   //Copy data
   FOR #i := 1 TO 9 DO
       #j := "HMI_OrderTable".StartRow + #i;
       "HMI_OrderTable".Index[#i] := #j;
       "HMI_OrderTable".OrderTable[#i] := #System.OrderTable[#j];
       //Color State
       IF "HMI_OrderTable".OrderTable[#i].Status = 'Queued' THEN
           "HMI_OrderTable".State[#i] := 1;
       ELSIF "HMI_OrderTable".OrderTable[#i].Status = 'Running' THEN
           "HMI_OrderTable".State[#i] := 2;
       ELSIF "HMI_OrderTable".OrderTable[#i].Status = 'Completed' THEN
           "HMI_OrderTable".State[#i] := 3;
       ELSIF "HMI_OrderTable".OrderTable[#i].Status = 'Error' THEN
           "HMI_OrderTable".State[#i] := 4;
       ELSIF "HMI_OrderTable".OrderTable[#i].Status = 'Paused' THEN
           "HMI_OrderTable".State[#i] := 5;
       ELSIF "HMI_OrderTable".OrderTable[#i].Status = 'Canceled' THEN
           "HMI_OrderTable".State[#i] := 6;
       ELSIF "HMI_OrderTable".OrderTable[#i].Status = 'Error\Cancel' THEN
           "HMI_OrderTable".State[#i] := 7;
       ELSE
           "HMI_OrderTable".State[#i] := 0;
       END_IF;
   END_FOR;

   IF NOT "HMI_OrderTable".PlacingNewOrder THEN
       "HMI_OrderTable".Device := 0;
   END_IF;

   //Error PopUp Window
   IF "HMI_OrderTable".PopUp_ErrorWindow_Active AND NOT "HMI_OrderTable".PlacingNewOrder THEN
       "HMI_OrderTable".OrderTable[0] := "HMI_OrderTable".OrderTable["HMI_OrderTable".PopUp_Index];
       IF "HMI_OrderTable".OrderTable[0].Status = 'Error' THEN
           "HMI_OrderTable".State[0] := 4;
       ELSIF "HMI_OrderTable".OrderTable[0].Status = 'Error\Cancel' THEN
           "HMI_OrderTable".State[0] := 7;
       ELSE
           "HMI_OrderTable".State[0] := 0;
       END_IF;
   ELSIF NOT "HMI_OrderTable".PopUp_ErrorWindow_Active AND NOT "HMI_OrderTable".PlacingNewOrder THEN
       "HMI_OrderTable".OrderTable[0] := #EmptyOrder;
   END_IF;

   REGION Testing area
       IF ("HMI_Box_Connected_1" = #System.Id OR ("HMI_Box_Connected_1" >= (#System.Id * 10) + 1 AND "HMI_Box_Connected_1" <= (#System.Id * 10) + 8)) OR
           ("HMI_Box_Connected_2" = #System.Id OR ("HMI_Box_Connected_1" >= (#System.Id * 10) + 1 AND "HMI_Box_Connected_1" <= (#System.Id * 10) + 8))
       THEN
           #System_Busy := TRUE;
       ELSE
           #System_Busy := FALSE;
           IF "Comissioning_Var" THEN
           //Visibilities
           //Running in auto mode
           IF #Auto_Test.Running AND NOT #Auto_Test.Manual AND NOT #Auto_Test.Pause THEN
               "OrderTable_HMI"."Start Test Visibility" := FALSE;
               "OrderTable_HMI"."Stop Test Visibility" := TRUE;
               "OrderTable_HMI"."Pause Test Visibility" := TRUE;
               "OrderTable_HMI"."Resume Visibility" := FALSE;
               "OrderTable_HMI"."Clear Table Visibility" := FALSE;
               "OrderTable_HMI"."Manual order Visibility" := FALSE;
               //Running and paused
           ELSIF #Auto_Test.Running AND #Auto_Test.Pause AND NOT #Auto_Test.Manual THEN
               "OrderTable_HMI"."Start Test Visibility" := FALSE;
               "OrderTable_HMI"."Stop Test Visibility" := TRUE;
               "OrderTable_HMI"."Pause Test Visibility" := FALSE;
               "OrderTable_HMI"."Resume Visibility" := TRUE;
               "OrderTable_HMI"."Clear Table Visibility" := FALSE;
               "OrderTable_HMI"."Manual order Visibility" := FALSE;
               //Running and Manual
           ELSIF #Auto_Test.Manual AND #Auto_Test.Running THEN
               "OrderTable_HMI"."Start Test Visibility" := FALSE;
               "OrderTable_HMI"."Stop Test Visibility" := FALSE;
               "OrderTable_HMI"."Pause Test Visibility" := FALSE;
               "OrderTable_HMI"."Resume Visibility" := FALSE;
               "OrderTable_HMI"."Clear Table Visibility" := FALSE;
               "OrderTable_HMI"."Manual order Visibility" := FALSE;
               //Manual and not running
           ELSIF #Auto_Test.Manual AND NOT #Auto_Test.Running THEN
               "OrderTable_HMI"."Start Test Visibility" := FALSE;
               "OrderTable_HMI"."Stop Test Visibility" := FALSE;
               "OrderTable_HMI"."Pause Test Visibility" := FALSE;
               "OrderTable_HMI"."Resume Visibility" := FALSE;
               "OrderTable_HMI"."Clear Table Visibility" := FALSE;
               "OrderTable_HMI"."Manual order Visibility" := TRUE;
               // not running, in automatic and no error
           ELSIF #Auto_Test.Automatic AND NOT #Auto_Test.Error AND #Auto_Test.State = 10 THEN
               "OrderTable_HMI"."Start Test Visibility" := TRUE;
               "OrderTable_HMI"."Stop Test Visibility" := FALSE;
               "OrderTable_HMI"."Pause Test Visibility" := FALSE;
               "OrderTable_HMI"."Resume Visibility" := FALSE;
               "OrderTable_HMI"."Clear Table Visibility" := TRUE;
               "OrderTable_HMI"."Manual order Visibility" := TRUE;
           ELSIF NOT #Auto_Test.Running THEN
               "OrderTable_HMI"."Clear Table Visibility" := TRUE;
               "OrderTable_HMI"."Manual order Visibility" := TRUE;
           END_IF;

           //PALLET TYPE VISIBILITY
           IF "OrderTable_HMI"."Pallet Type" = 1 THEN //CHEP
               "OrderTable_HMI"."Tower 1 Visibility" := FALSE;
               "OrderTable_HMI"."Tower 2 Visibility" := FALSE;
               "OrderTable_HMI"."Extractor Visibility" := FALSE;
           ELSIF "OrderTable_HMI"."Pallet Type" = 2 THEN //EURO
               "OrderTable_HMI"."Tower 1 Visibility" := TRUE;
               "OrderTable_HMI"."Tower 2 Visibility" := TRUE;
               "OrderTable_HMI"."Extractor Visibility" := TRUE;
           END_IF;

           IF #Auto_Test.Manual THEN
               "OrderTable_HMI"."Tower Visibility" := TRUE;
               "OrderTable_HMI"."Level Visibility" := TRUE;
               "OrderTable_HMI"."ToExtractor Visibility" := TRUE;
               "OrderTable_HMI".Auto_Settings_Visibility := FALSE;
               IF #Auto_Test.Level <> 0 AND NOT #Auto_Test.Running THEN
                   "OrderTable_HMI"."Send VTD Order Visibility" := TRUE;
               END_IF;
               IF (("OrderTable_HMI"."Pallet Type" = 1) OR
                   ("OrderTable_HMI"."Pallet Type" = 2 AND "OrderTable_HMI".Tower = 1 AND "OrderTable_HMI"."Tower 1 Pallet Alignment" <> 0 AND "OrderTable_HMI".Transfer_From_To = 2) OR
                   ("OrderTable_HMI"."Pallet Type" = 2 AND "OrderTable_HMI".Tower = 2 AND "OrderTable_HMI"."Tower 1 Pallet Alignment" <> 0 AND "OrderTable_HMI".Transfer_From_To = 2) OR
                   ("OrderTable_HMI"."Pallet Type" = 2 AND "OrderTable_HMI"."Extractor Pallet Alignment" <> 0 AND "OrderTable_HMI".Transfer_From_To = 1))
                   AND
                   "OrderTable_HMI".Tower <> 0 AND "OrderTable_HMI".Transfer_From_To <> 0 AND NOT #Auto_Test.Running THEN
                   "OrderTable_HMI"."Send CNV Order Visibility" := TRUE;
               ELSE
                   "OrderTable_HMI"."Send CNV Order Visibility" := FALSE;
               END_IF;
           ELSE
               "OrderTable_HMI"."Tower Visibility" := FALSE;
               "OrderTable_HMI"."Level Visibility" := FALSE;
               "OrderTable_HMI"."ToExtractor Visibility" := FALSE;
               "OrderTable_HMI".Auto_Settings_Visibility := TRUE;
               "OrderTable_HMI"."Send VTD Order Visibility" := FALSE;
               "OrderTable_HMI"."Send CNV Order Visibility" := FALSE;
           END_IF;

           "OrderTable_HMI"."Pallet Type Visibility" := TRUE;
       ELSE
           "OrderTable_HMI"."Tower Visibility" := FALSE;
           "OrderTable_HMI"."Level Visibility" := FALSE;
           "OrderTable_HMI"."ToExtractor Visibility" := FALSE;
           "OrderTable_HMI".Auto_Settings_Visibility := FALSE;
           "OrderTable_HMI"."Send VTD Order Visibility" := FALSE;
           "OrderTable_HMI"."Send CNV Order Visibility" := FALSE;
           "OrderTable_HMI"."Pallet Type Visibility" := FALSE;
           "OrderTable_HMI"."Clear Table Visibility" := TRUE;
           "OrderTable_HMI"."Manual order Visibility" := FALSE;
       END_IF;

           //Buttons actions
           //START
           IF "OrderTable_HMI".Start THEN
               #Auto_Test.Start := TRUE;
           END_IF;

           //PAUSE
           IF "OrderTable_HMI".Pause THEN
               #Auto_Test.Pause := TRUE;
           END_IF;

           //STOP
           IF "OrderTable_HMI".Stop THEN
               #Auto_Test.Stop := TRUE;
           ELSE
               #Auto_Test.Stop := FALSE;
           END_IF;

           //RESUME
           IF "OrderTable_HMI".Resume THEN
               #Auto_Test.Pause := FALSE;
           END_IF;

           //MANUAL
           #Auto_Test.Manual := "OrderTable_HMI"."Manual order";

           //SEND VTD ORDER
           "R_Send_VTD_Order"(CLK := "OrderTable_HMI"."Send VTD Order");
           IF "R_Send_VTD_Order".Q THEN
               #Auto_Test.Send_VTD_Order := TRUE;
           END_IF;

           //SEND CNV ORDER
           "R_Send_CNV_Order"(CLK := "OrderTable_HMI"."Send CNV Order");
           IF "R_Send_CNV_Order".Q THEN
               #Auto_Test.Send_CNV_Order := TRUE;
           END_IF;

           //TEST SETTINGS
           //PALLET TYPE
           IF "OrderTable_HMI"."Pallet Type" = 1 THEN
               #Auto_Test."Pallet Type" := 'C';
           ELSIF "OrderTable_HMI"."Pallet Type" = 2 THEN
               #Auto_Test."Pallet Type" := 'E';
           ELSE
               #Auto_Test."Pallet Type" := ' ';
           END_IF;

           //PALLET ALIGNMENT TOWER 1
           IF "OrderTable_HMI"."Tower 1 Pallet Alignment" = 1 AND
               (("OrderTable_HMI".Transfer_From_To = 2 AND #Auto_Test.Manual) OR NOT #Auto_Test.Manual) THEN
               #Auto_Test."Tower 1 Pallet Alignment" := 'R';
               #Auto_Test.Pallet_Allignment := 'R';
           ELSIF "OrderTable_HMI"."Tower 1 Pallet Alignment" = 2 AND
               (("OrderTable_HMI".Transfer_From_To = 2 AND #Auto_Test.Manual) OR NOT #Auto_Test.Manual) THEN
               #Auto_Test."Tower 1 Pallet Alignment" := 'L';
               #Auto_Test.Pallet_Allignment := 'L';
           END_IF;

           //PALLET ALIGNMENT ECONVEYOR
           IF "OrderTable_HMI"."Extractor Pallet Alignment" = 1 AND
               (("OrderTable_HMI".Transfer_From_To = 1 AND #Auto_Test.Manual) OR NOT #Auto_Test.Manual) THEN
               #Auto_Test."Extractor Pallet Alignment" := 'R';
               #Auto_Test.Pallet_Allignment := 'R';
           ELSIF "OrderTable_HMI"."Extractor Pallet Alignment" = 2 AND
               (("OrderTable_HMI".Transfer_From_To = 1 AND #Auto_Test.Manual) OR NOT #Auto_Test.Manual) THEN
               #Auto_Test."Extractor Pallet Alignment" := 'L';
               #Auto_Test.Pallet_Allignment := 'L';
           ELSIF "OrderTable_HMI"."Extractor Pallet Alignment" = 3 AND
               (("OrderTable_HMI".Transfer_From_To = 1 AND #Auto_Test.Manual) OR NOT #Auto_Test.Manual) THEN
               #Auto_Test."Extractor Pallet Alignment" := 'C';
               #Auto_Test.Pallet_Allignment := 'C';
           END_IF;

           //AUTOMATIC SETTING FOR BUTTON TRANSFER FROM_TO
           IF NOT "Control_DB".VTD_Sys[#Sys].Running AND "Control_DB".VTD_Sys[#Sys].Current_Level <> 0 THEN
               IF #Auto_Test.Tower = 1 AND "HMI_DB".ScreenNo_Main = 9 THEN
                   //CNV 1
                   IF "Control_DB".ECnv_Sys[#Sys].Cnv_Occupied AND NOT "Control_DB".LCnv_Sys[#Sys].Cnv_Level["Control_DB".VTD_Sys[#Sys].Current_Level].Cnv1.Cnv_Occupied AND
                       NOT "Control_DB".ECnv_Sys[#Sys].Running AND NOT "Control_DB".LCnv_Sys[#Sys].Cnv_Level["Control_DB".VTD_Sys[#Sys].Current_Level].Cnv1.Running THEN
                       #Auto_Test.Transfer_From_To := "OrderTable_HMI".Transfer_From_To := 2;//to buffer
                   ELSIF NOT "Control_DB".ECnv_Sys[#Sys].Cnv_Occupied AND "Control_DB".LCnv_Sys[#Sys].Cnv_Level["Control_DB".VTD_Sys[#Sys].Current_Level].Cnv1.Cnv_Occupied AND
                       NOT "Control_DB".ECnv_Sys[#Sys].Running AND NOT "Control_DB".LCnv_Sys[#Sys].Cnv_Level["Control_DB".VTD_Sys[#Sys].Current_Level].Cnv1.Running THEN
                       #Auto_Test.Transfer_From_To := "OrderTable_HMI".Transfer_From_To := 1;//to extractor
                   ELSE
                       #Auto_Test.Transfer_From_To := "OrderTable_HMI".Transfer_From_To;
                   END_IF;
                   //CNV 2
               ELSIF #Auto_Test.Tower = 2 AND "HMI_DB".ScreenNo_Main = 9 THEN   //CNV 2
                   IF "Control_DB".ECnv_Sys[#Sys].Cnv_Occupied AND NOT "Control_DB".LCnv_Sys[#Sys].Cnv_Level["Control_DB".VTD_Sys[#Sys].Current_Level].Cnv2.Cnv_Occupied AND
                       NOT "Control_DB".ECnv_Sys[#Sys].Running AND NOT "Control_DB".LCnv_Sys[#Sys].Cnv_Level["Control_DB".VTD_Sys[#Sys].Current_Level].Cnv2.Running THEN
                       #Auto_Test.Transfer_From_To := "OrderTable_HMI".Transfer_From_To := 2;
                   ELSIF NOT "Control_DB".ECnv_Sys[#Sys].Cnv_Occupied AND "Control_DB".LCnv_Sys[#Sys].Cnv_Level["Control_DB".VTD_Sys[#Sys].Current_Level].Cnv2.Cnv_Occupied AND
                       NOT "Control_DB".ECnv_Sys[#Sys].Running AND NOT "Control_DB".LCnv_Sys[#Sys].Cnv_Level["Control_DB".VTD_Sys[#Sys].Current_Level].Cnv2.Running THEN
                       #Auto_Test.Transfer_From_To := "OrderTable_HMI".Transfer_From_To := 1;
                   ELSE
                       #Auto_Test.Transfer_From_To := "OrderTable_HMI".Transfer_From_To;
                   END_IF;
               END_IF;
           END_IF;

           //LEVELS AND CYCLES
           #Auto_Test."From level" := "OrderTable_HMI"."From level";
           #Auto_Test."To level" := "OrderTable_HMI"."To level";
           #Auto_Test."Testing Time" := "OrderTable_HMI"."Testing Time";
           #Auto_Test."Numer of cycles" := "OrderTable_HMI"."Numer of cycles";
           #Auto_Test.Level := "OrderTable_HMI".Level;
           #Auto_Test.Tower := "OrderTable_HMI".Tower;
           "OrderTable_HMI"."Time Running" := DINT_TO_UINT(TIME_TO_DINT(#Auto_Test.Time_Runnng) / 60000);
           "OrderTable_HMI".Actual_Cycle := UINT_TO_BYTE(#Auto_Test.N_Cycles);
       END_IF;
   END_REGION ;
END_FUNCTION

FUNCTION_BLOCK "F_Lock_FB"   // FB24, F_FBD
{ S7_Optimized_Access := 'TRUE' }
VERSION : 0.1
// stored: AutoNumber true, IsIECCheckEnabled false, UDAEnableTagReadback false
   VAR_INPUT
      Lock_Closed_CH1 { ExternalAccessible := 'False'; ExternalVisible := 'False'; ExternalWritable := 'False'} : Bool;
      Lock_Closed_CH2 { ExternalAccessible := 'False'; ExternalVisible := 'False'; ExternalWritable := 'False'} : Bool;
      EStop_CH1 { ExternalAccessible := 'False'; ExternalVisible := 'False'; ExternalWritable := 'False'} : Bool;
      EStop_CH2 { ExternalAccessible := 'False'; ExternalVisible := 'False'; ExternalWritable := 'False'} : Bool;
      ACK { ExternalAccessible := 'False'; ExternalVisible := 'False'; ExternalWritable := 'False'} : Bool;
   END_VAR
   VAR_OUTPUT
      Lock_Reset_Input1 { ExternalAccessible := 'False'; ExternalVisible := 'False'; ExternalWritable := 'False'} : Bool;
      Lock_Reset_Input2 { ExternalAccessible := 'False'; ExternalVisible := 'False'; ExternalWritable := 'False'} : Bool;
      Lock_Reset_Input3 { ExternalAccessible := 'False'; ExternalVisible := 'False'; ExternalWritable := 'False'} : Bool;
      Lock_Reset_Input4 { ExternalAccessible := 'False'; ExternalVisible := 'False'; ExternalWritable := 'False'} : Bool;
      EStop_Lock_OK : Bool;
      Lock_Secured_OK : Bool;
   END_VAR
   VAR
      GUARD_SWITCH : ESTOP1;
      ESTOP : ESTOP1;
   END_VAR
BEGIN

REGION Network 1: GUARD SWITCH
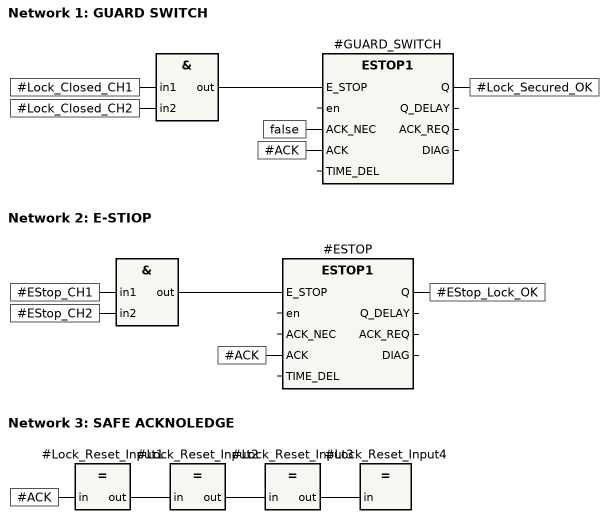
   #GUARD_SWITCH(E_STOP := #Lock_Closed_CH1 AND #Lock_Closed_CH2,   // ESTOP1
                 ACK_NEC := false,
                 ACK := #ACK,
                 Q => #Lock_Secured_OK);
END_REGION

REGION Network 2: E-STIOP
   #ESTOP(E_STOP := #EStop_CH1 AND #EStop_CH2, ACK := #ACK, Q => #EStop_Lock_OK);   // ESTOP1
END_REGION

REGION Network 3: SAFE ACKNOLEDGE
   #Lock_Reset_Input1 := #ACK;
   #Lock_Reset_Input2 := #ACK;
   #Lock_Reset_Input3 := #ACK;
   #Lock_Reset_Input4 := #ACK;
END_REGION
END_FUNCTION_BLOCK

FUNCTION "Feed_BCNV_Cnv1(1)" : Void   // FC54, SCL
{ S7_Optimized_Access := 'TRUE' }
VERSION : 0.1
// stored: AutoNumber true, IsIECCheckEnabled false, SetENOAutomatically false, UDAEnableTagReadback false
   VAR_INPUT
      System_No : UInt;
      Level : UInt;
      Light_Guard_IO : Bool;
   END_VAR
   VAR_OUTPUT
      Light_Guard_Bypass : Bool;
   END_VAR
   VAR_IN_OUT
      System_Busy : Bool;
   END_VAR
BEGIN
   //Sensors
   "HMI_CNV_Left(1)" := "Control_DB".LCnv_Sys[#System_No].Cnv_Level[#Level].Cnv1.Inputs.Left;
   "HMI_CNV_Lpd1(1)" := "Control_DB".LCnv_Sys[#System_No].Cnv_Level[#Level].Cnv1.Inputs.Lpd1;
   "HMI_CNV_Lpd2(1)" := "Control_DB".LCnv_Sys[#System_No].Cnv_Level[#Level].Cnv1.Inputs.Lpd2;
   "HMI_CNV_Right(1)" := "Control_DB".LCnv_Sys[#System_No].Cnv_Level[#Level].Cnv1.Inputs.Right;
   "HMI_CNV_Rpd1(1)" := "Control_DB".LCnv_Sys[#System_No].Cnv_Level[#Level].Cnv1.Inputs.Rpd1;
   "HMI_CNV_Rpd2(1)" := "Control_DB".LCnv_Sys[#System_No].Cnv_Level[#Level].Cnv1.Inputs.Rpd2;
   "HMI_CNV_Sdetect1(1)" := "Control_DB".LCnv_Sys[#System_No].Cnv_Level[#Level].Cnv1.Inputs.Sdetect1;
   "HMI_CNV_Sdetect2(1)" := "Control_DB".LCnv_Sys[#System_No].Cnv_Level[#Level].Cnv1.Inputs.Sdetect2;
   "HMI_CNV_SftyPinUp(1)" := "Control_DB".LCnv_Sys[#System_No].Cnv_Level[#Level].Cnv1.Safety_Stop_Cnrl.Inputs.DP_Extended;
   "HMI_CNV_SftyPinDown(1)" := "Control_DB".LCnv_Sys[#System_No].Cnv_Level[#Level].Cnv1.Safety_Stop_Cnrl.Inputs.DP_Retracted;
   "HMI_Light_Guard" := #System_No <= 3 AND #Level = 1 AND "HMI_DB".Username = 'admin'; //To show the button
   IF "Control_DB".LCnv_Sys[#System_No].Cnv_Level[#Level].Cnv1.Safety_Stop_Cnrl.Inputs.DP_Extended AND
       NOT "Control_DB".LCnv_Sys[#System_No].Cnv_Level[#Level].Cnv1.Safety_Stop_Cnrl.Inputs.DP_Retracted THEN
       "UpDown(1)" := 1;
   ELSIF NOT "Control_DB".LCnv_Sys[#System_No].Cnv_Level[#Level].Cnv1.Safety_Stop_Cnrl.Inputs.DP_Extended AND
       "Control_DB".LCnv_Sys[#System_No].Cnv_Level[#Level].Cnv1.Safety_Stop_Cnrl.Inputs.DP_Retracted THEN
       "UpDown(1)" := 2;
   ELSE
       "UpDown(1)" := 0;
   END_IF;

   //Status
   "Mode_HMI(1)" := "Control_DB".LCnv_Sys[#System_No].Cnv_Level[#Level].Cnv1.Mode;
   "Enabled_HMI(1)" := "Control_DB".LCnv_Sys[#System_No].Cnv_Level[#Level].Cnv1.Enabled;
   "Error_HMI(1)" := "Control_DB".LCnv_Sys[#System_No].Cnv_Level[#Level].Cnv1.Error;
   "Warning_HMI(1)" := "Control_DB".LCnv_Sys[#System_No].Cnv_Level[#Level].Cnv1.Warning;
   "Stopped_HMI(1)" := "Control_DB".LCnv_Sys[#System_No].Cnv_Level[#Level].Cnv1.Stopped;
   "Running_HMI(1)" := "Control_DB".LCnv_Sys[#System_No].Cnv_Level[#Level].Cnv1.Running;
   "Ready_For_Task_HMI(1)" := "Control_DB".LCnv_Sys[#System_No].Cnv_Level[#Level].Cnv1.Ready_For_Task;
   "Cnv_Occupied_HMI(1)" := "Control_DB".LCnv_Sys[#System_No].Cnv_Level[#Level].Cnv1.Cnv_Occupied;
   "Shuttle_in_place_HMI(1)" := "Control_DB".LCnv_Sys[#System_No].Cnv_Level[#Level].Cnv1.Shuttle_In_Place;
   "Current_Task_Type_HMI(1)" := "Control_DB".LCnv_Sys[#System_No].Cnv_Level[#Level].Cnv1.Current_Task_Type;
   "Current_Task_ID_HMI(1)" := "Control_DB".LCnv_Sys[#System_No].Cnv_Level[#Level].Cnv1.Current_Task_ID;
   "SM_State_HMI(1)" := "Control_DB".LCnv_Sys[#System_No].Cnv_Level[#Level].Cnv1.SM_State;
   "Pallet_Type_HMI(1)" := "Control_DB".LCnv_Sys[#System_No].Cnv_Level[#Level].Cnv1.Pallet_Type;
   IF "Control_DB".LCnv_Sys[#System_No].Cnv_Level[#Level].Cnv1.Motor.Forward THEN
       "Motor_Direction_HMI(1)" := 1;
   ELSIF "Control_DB".LCnv_Sys[#System_No].Cnv_Level[#Level].Cnv1.Motor.Reverse THEN
       "Motor_Direction_HMI(1)" := 2;
   ELSE
       "Motor_Direction_HMI(1)" := 0;
   END_IF;
   "Motor_Speed_Requested_HMI(1)" := "Control_DB".LCnv_Sys[#System_No].Cnv_Level[#Level].Cnv1.Motor.Speed;
   "Motor_Speed_Actual_HMI(1)" := "Control_DB".LCnv_Sys[#System_No].Cnv_Level[#Level].Cnv1.Motor.Speed_Actual;
   "CNV_Motor_Ready(1)" := "Control_DB".LCnv_Sys[#System_No].Cnv_Level[#Level].Cnv1.Motor.Ready;
   "CNV_Motor_Current_Actual_HMI(1)" := "Control_DB".LCnv_Sys[#System_No].Cnv_Level[#Level].Cnv1.Motor.Actual_Current;
   "CNV_Motor_Actual_Torque(1)" := "Control_DB".LCnv_Sys[#System_No].Cnv_Level[#Level].Cnv1.Motor.Actual_Torque;
   "Transfer_To_ID_HMI(1)" := "Control_DB".LCnv_Sys[#System_No].Cnv_Level[#Level].Cnv1.Instruction.Transfer_To_ID;
   "Transfer_From_ID_HMI(1)" := "Control_DB".LCnv_Sys[#System_No].Cnv_Level[#Level].Cnv1.Instruction.Transfer_From_ID;

   IF "Control_DB".LCnv_Sys[#System_No].Cnv_Level[#Level].Cnv1.Motor.Error THEN
       "CNV_Motor_Status_HMI(1)" := 2;
   ELSIF "Control_DB".LCnv_Sys[#System_No].Cnv_Level[#Level].Cnv1.Motor.Enabled THEN
       "CNV_Motor_Status_HMI(1)" := 1;
   ELSIF NOT "Control_DB".LCnv_Sys[#System_No].Cnv_Level[#Level].Cnv1.Motor.Enabled THEN
       "CNV_Motor_Status_HMI(1)" := 0;
   END_IF;

   //Instructions
   IF ("HMI_Box_Connected_1" = #System_No OR ("HMI_Box_Connected_1" >= (#System_No * 10) + 1 AND "HMI_Box_Connected_1" <= (#System_No * 10) + 8)) OR
       ("HMI_Box_Connected_2" = #System_No OR ("HMI_Box_Connected_1" >= (#System_No * 10) + 1 AND "HMI_Box_Connected_1" <= (#System_No * 10) + 8))
   THEN
       #System_Busy := TRUE;
   ELSE
       #System_Busy := FALSE;
       "Control_DB".LCnv_Sys[#System_No].Cnv_Level[#Level].Cnv1.Instruction.Stop := "Stop_HMI(1)";
       "Control_DB".LCnv_Sys[#System_No].Cnv_Level[#Level].Cnv1.Instruction.Execute := "Manual_Fwd_HMI(1)" OR "Manual_Bwd_HMI(1)";
       IF "BT_Confirmation_HMI" THEN
           "Control_DB".VTD_Sys[#System_No].Instruction.Mode_Change :=
           "Control_DB".ECnv_Sys[#System_No].Instruction.Mode_Change :=
           "Control_DB".LCnv_Sys[#System_No].Cnv_Level[1].Cnv1.Instruction.Mode_Change :=
           "Control_DB".LCnv_Sys[#System_No].Cnv_Level[2].Cnv1.Instruction.Mode_Change :=
           "Control_DB".LCnv_Sys[#System_No].Cnv_Level[3].Cnv1.Instruction.Mode_Change :=
           "Control_DB".LCnv_Sys[#System_No].Cnv_Level[4].Cnv1.Instruction.Mode_Change :=
           "Control_DB".LCnv_Sys[#System_No].Cnv_Level[5].Cnv1.Instruction.Mode_Change :=
           "Control_DB".LCnv_Sys[#System_No].Cnv_Level[6].Cnv1.Instruction.Mode_Change :=
           "Control_DB".LCnv_Sys[#System_No].Cnv_Level[7].Cnv1.Instruction.Mode_Change :=
           "Control_DB".LCnv_Sys[#System_No].Cnv_Level[8].Cnv1.Instruction.Mode_Change :=
           "Control_DB".LCnv_Sys[#System_No].Cnv_Level[1].Cnv2.Instruction.Mode_Change :=
           "Control_DB".LCnv_Sys[#System_No].Cnv_Level[2].Cnv2.Instruction.Mode_Change :=
           "Control_DB".LCnv_Sys[#System_No].Cnv_Level[3].Cnv2.Instruction.Mode_Change :=
           "Control_DB".LCnv_Sys[#System_No].Cnv_Level[4].Cnv2.Instruction.Mode_Change :=
           "Control_DB".LCnv_Sys[#System_No].Cnv_Level[5].Cnv2.Instruction.Mode_Change :=
           "Control_DB".LCnv_Sys[#System_No].Cnv_Level[6].Cnv2.Instruction.Mode_Change :=
           "Control_DB".LCnv_Sys[#System_No].Cnv_Level[7].Cnv2.Instruction.Mode_Change :=
           "Control_DB".LCnv_Sys[#System_No].Cnv_Level[8].Cnv2.Instruction.Mode_Change := "Mode_Change_HMI(1)";
           "Mode_Change_HMI" := "Mode_Change_HMI(1)";
           "BT_Confirmation_HMI" := FALSE;
       END_IF;

       "Control_DB".LCnv_Sys[#System_No].Cnv_Level[#Level].Cnv1.Instruction.Enable := "Enable_HMI(1)";
       IF "Control_DB".LCnv_Sys[#System_No].Cnv_Level[#Level].Cnv1.Mode <> 1 THEN
           "HMI_Light_Guard_Bypass" := FALSE;
       ELSIF "HMI_Light_Guard_Bypass" AND "Control_DB".LCnv_Sys[#System_No].Cnv_Level[1].Cnv1.Error THEN
           #Light_Guard_Bypass := TRUE;
       ELSIF NOT "Control_DB".LCnv_Sys[#System_No].Cnv_Level[1].Cnv1.Running AND NOT "Control_DB".LCnv_Sys[#System_No].Cnv_Level[1].Cnv1.Error AND #Light_Guard_IO THEN //Not Running and No error and light guard free
           #Light_Guard_Bypass := FALSE; //Cancel bypass
       END_IF;

       IF "Control_DB".LCnv_Sys[#System_No].Cnv_Level[#Level].Cnv1.Mode <> 3 THEN
           "Control_DB".LCnv_Sys[#System_No].Cnv_Level[#Level].Cnv1.Instruction.Foward := "Manual_Fwd_HMI(1)";
           "Control_DB".LCnv_Sys[#System_No].Cnv_Level[#Level].Cnv1.Instruction.Backward := "Manual_Bwd_HMI(1)";
           "Control_DB".LCnv_Sys[#System_No].Cnv_Level[#Level].Cnv1.Instruction.Start_Transfer := "Start_Transfer_HMI(1)";
           IF "Control_DB".LCnv_Sys[#System_No].Cnv_Level[#Level].Cnv1.Mode = 1 THEN
               "Control_DB".LCnv_Sys[#System_No].Cnv_Level[#Level].Cnv1.Instruction.Start_Transfer_Backward := "Transfer_Backward(1)";
           END_IF;
           "Control_DB".LCnv_Sys[#System_No].Cnv_Level[#Level].Cnv1.Safety_Stop_Cnrl.Instruction.Manual_Extend := "Manual_Sfty_Stopper_Up(1)";
           "Control_DB".LCnv_Sys[#System_No].Cnv_Level[#Level].Cnv1.Safety_Stop_Cnrl.Instruction.Manual_Retract := "Manual_Sfty_Stopper_Down(1)";
           "Control_DB".LCnv_Sys[#System_No].Cnv_Level[#Level].Cnv1.Instruction.Task_ID := "Task_ID_HMI(1)";
           "Control_DB".LCnv_Sys[#System_No].Cnv_Level[#Level].Cnv1.Instruction.Pallet_Align_Left := "Pallet_Align_Left_HMI(1)";
           "Control_DB".LCnv_Sys[#System_No].Cnv_Level[#Level].Cnv1.Instruction.Pallet_Align_Right := "Pallet_Align_Right_HMI(1)";
           IF "Mode_Change_HMI(1)" <> 2 THEN
               "Control_DB".LCnv_Sys[#System_No].Cnv_Level[#Level].Cnv1.Instruction.Pallet_Allignment := "Pallet_Allignment_HMI(1)" := FALSE;
           ELSE
               "Control_DB".LCnv_Sys[#System_No].Cnv_Level[#Level].Cnv1.Instruction.Pallet_Allignment := "Pallet_Allignment_HMI(1)";
           END_IF;
           IF "CNV_HMI".In_Out[#System_No] THEN // 0 = ECNV RECEIVE, 1 = ECONV SEND
               "Control_DB".LCnv_Sys[#System_No].Cnv_Level[#Level].Cnv1.Instruction.Transfer_To_ID := 0;
               "Control_DB".LCnv_Sys[#System_No].Cnv_Level[#Level].Cnv1.Instruction.Transfer_From_ID := DINT#120000 + (#Level * 100) + #System_No;
           ELSE
               "Control_DB".LCnv_Sys[#System_No].Cnv_Level[#Level].Cnv1.Instruction.Transfer_To_ID := DINT#120000 + (#Level * 100) + #System_No;
               "Control_DB".LCnv_Sys[#System_No].Cnv_Level[#Level].Cnv1.Instruction.Transfer_From_ID := 0;
           END_IF;
       END_IF;

       "Control_DB".LCnv_Sys[#System_No].Cnv_Level[#Level].Cnv1.Instruction.Reset :=
       "Reset_HMI(1)" OR "Reset_All" OR
       "CNV_HMI"."Reset(1)"[1] OR "Screen_DB_1".Reset_All[1] OR
       "CNV_HMI"."Reset(1)"[2] OR "Screen_DB_1".Reset_All[2];
   END_IF;
END_FUNCTION

FUNCTION "Feed_BCNV_Cnv1(1)_1" : Void   // FC56, SCL
{ S7_Optimized_Access := 'TRUE' }
VERSION : 0.1
// stored: AutoNumber true, IsIECCheckEnabled false, SetENOAutomatically false, UDAEnableTagReadback false
   VAR_INPUT
      HMI_No : UInt;
      System_No : UInt;
      Level : UInt;
      Light_Guard_IO : Bool;
   END_VAR
   VAR_OUTPUT
      Light_Guard_Bypass : Bool;
   END_VAR
BEGIN
   //Sensors
   "CNV_HMI"."Left(1)"[#HMI_No] := "Control_DB".LCnv_Sys[#System_No].Cnv_Level[#Level].Cnv1.Inputs.Left;
   "CNV_HMI"."Lpd1(1)"[#HMI_No] := "Control_DB".LCnv_Sys[#System_No].Cnv_Level[#Level].Cnv1.Inputs.Lpd1;
   "CNV_HMI"."Lpd2(1)"[#HMI_No] := "Control_DB".LCnv_Sys[#System_No].Cnv_Level[#Level].Cnv1.Inputs.Lpd2;
   "CNV_HMI"."Right(1)"[#HMI_No] := "Control_DB".LCnv_Sys[#System_No].Cnv_Level[#Level].Cnv1.Inputs.Right;
   "CNV_HMI"."Rpd1(1)"[#HMI_No] := "Control_DB".LCnv_Sys[#System_No].Cnv_Level[#Level].Cnv1.Inputs.Rpd1;
   "CNV_HMI"."Rpd2(1)"[#HMI_No] := "Control_DB".LCnv_Sys[#System_No].Cnv_Level[#Level].Cnv1.Inputs.Rpd2;
   "CNV_HMI"."Sdetect1(1)"[#HMI_No] := "Control_DB".LCnv_Sys[#System_No].Cnv_Level[#Level].Cnv1.Inputs.Sdetect1;
   "CNV_HMI"."Sdetect2(1)"[#HMI_No] := "Control_DB".LCnv_Sys[#System_No].Cnv_Level[#Level].Cnv1.Inputs.Sdetect2;
   "HMI_Light_Guard" := #Level = 1; //To show the button
   IF "Control_DB".LCnv_Sys[#System_No].Cnv_Level[#Level].Cnv1.Safety_Stop_Cnrl.Inputs.DP_Extended AND
       NOT "Control_DB".LCnv_Sys[#System_No].Cnv_Level[#Level].Cnv1.Safety_Stop_Cnrl.Inputs.DP_Retracted THEN
       "CNV_HMI"."UpDown(1)"[#HMI_No] := 1;
   ELSIF NOT "Control_DB".LCnv_Sys[#System_No].Cnv_Level[#Level].Cnv1.Safety_Stop_Cnrl.Inputs.DP_Extended AND
       "Control_DB".LCnv_Sys[#System_No].Cnv_Level[#Level].Cnv1.Safety_Stop_Cnrl.Inputs.DP_Retracted THEN
       "CNV_HMI"."UpDown(1)"[#HMI_No] := 2;
   ELSE
       "CNV_HMI"."UpDown(1)"[#HMI_No] := 0;
   END_IF;

   //Status
   "CNV_HMI"."Mode(1)"[#HMI_No] := "Control_DB".LCnv_Sys[#System_No].Cnv_Level[#Level].Cnv1.Mode;
   "CNV_HMI"."Enabled(1)"[#HMI_No] := "Control_DB".LCnv_Sys[#System_No].Cnv_Level[#Level].Cnv1.Enabled;
   "CNV_HMI"."Error(1)"[#HMI_No] := "Control_DB".LCnv_Sys[#System_No].Cnv_Level[#Level].Cnv1.Error;
   "CNV_HMI"."Warning(1)"[#HMI_No] := "Control_DB".LCnv_Sys[#System_No].Cnv_Level[#Level].Cnv1.Warning;
   "CNV_HMI"."Stopped(1)"[#HMI_No] := "Control_DB".LCnv_Sys[#System_No].Cnv_Level[#Level].Cnv1.Stopped;
   "CNV_HMI"."Running(1)"[#HMI_No] := "Control_DB".LCnv_Sys[#System_No].Cnv_Level[#Level].Cnv1.Running;
   "CNV_HMI"."Ready_For_Task(1)"[#HMI_No] := "Control_DB".LCnv_Sys[#System_No].Cnv_Level[#Level].Cnv1.Ready_For_Task;
   "CNV_HMI"."Occupied(1)"[#HMI_No] := "Control_DB".LCnv_Sys[#System_No].Cnv_Level[#Level].Cnv1.Cnv_Occupied;
   "CNV_HMI"."Shuttle_in_place(1)"[#HMI_No] := "Control_DB".LCnv_Sys[#System_No].Cnv_Level[#Level].Cnv1.Shuttle_In_Place;
   "CNV_HMI"."Current_Task_Type(1)"[#HMI_No] := "Control_DB".LCnv_Sys[#System_No].Cnv_Level[#Level].Cnv1.Current_Task_Type;
   "CNV_HMI"."Task_ID(1)"[#HMI_No] := "Control_DB".LCnv_Sys[#System_No].Cnv_Level[#Level].Cnv1.Current_Task_ID;
   "CNV_HMI"."SM_State(1)"[#HMI_No] := "Control_DB".LCnv_Sys[#System_No].Cnv_Level[#Level].Cnv1.SM_State;
   "CNV_HMI"."Pallet_Type(1)"[#HMI_No] := "Control_DB".LCnv_Sys[#System_No].Cnv_Level[#Level].Cnv1.Pallet_Type;
   IF "Control_DB".LCnv_Sys[#System_No].Cnv_Level[#Level].Cnv1.Motor.Forward THEN
       "CNV_HMI"."Motor_Direction(1)"[#HMI_No] := 1;
   ELSIF "Control_DB".LCnv_Sys[#System_No].Cnv_Level[#Level].Cnv1.Motor.Reverse THEN
       "CNV_HMI"."Motor_Direction(1)"[#HMI_No] := 2;
   ELSE
       "CNV_HMI"."Motor_Direction(1)"[#HMI_No] := 0;
   END_IF;
   "CNV_HMI"."Motor_Speed_Requested(1)"[#HMI_No] := "Control_DB".LCnv_Sys[#System_No].Cnv_Level[#Level].Cnv1.Motor.Speed;
   "CNV_HMI"."Motor_Speed_Actual(1)"[#HMI_No] := "Control_DB".LCnv_Sys[#System_No].Cnv_Level[#Level].Cnv1.Motor.Speed_Actual;
   "CNV_HMI"."Motor_Ready(1)"[#HMI_No] := "Control_DB".LCnv_Sys[#System_No].Cnv_Level[#Level].Cnv1.Motor.Ready;
   "CNV_HMI"."Motor_Current_Actual(1)"[#HMI_No] := "Control_DB".LCnv_Sys[#System_No].Cnv_Level[#Level].Cnv1.Motor.Actual_Current;
   "CNV_HMI"."Motor_Actual_Torque(1)"[#HMI_No] := "Control_DB".LCnv_Sys[#System_No].Cnv_Level[#Level].Cnv1.Motor.Actual_Torque;
   "CNV_HMI"."Transfer_To_ID(1)"[#HMI_No] := "Control_DB".LCnv_Sys[#System_No].Cnv_Level[#Level].Cnv1.Instruction.Transfer_To_ID;
   "CNV_HMI"."Transfer_From_ID(1)"[#HMI_No] := "Control_DB".LCnv_Sys[#System_No].Cnv_Level[#Level].Cnv1.Instruction.Transfer_From_ID;

   IF "Control_DB".LCnv_Sys[#System_No].Cnv_Level[#Level].Cnv1.Motor.Error THEN
       "CNV_HMI"."Motor_Status(1)"[#HMI_No] := 2;
   ELSIF "Control_DB".LCnv_Sys[#System_No].Cnv_Level[#Level].Cnv1.Motor.Enabled THEN
       "CNV_HMI"."Motor_Status(1)"[#HMI_No] := 1;
   ELSIF NOT "Control_DB".LCnv_Sys[#System_No].Cnv_Level[#Level].Cnv1.Motor.Enabled THEN
       "CNV_HMI"."Motor_Status(1)"[#HMI_No] := 0;
   END_IF;

   //Instructions
   "Control_DB".LCnv_Sys[#System_No].Cnv_Level[#Level].Cnv1.Instruction.Stop := "CNV_HMI"."Stop(1)"[#HMI_No];
   "Control_DB".LCnv_Sys[#System_No].Cnv_Level[#Level].Cnv1.Instruction.Execute := "CNV_HMI"."Manual_Fwd(1)"[#HMI_No] OR "CNV_HMI"."Manual_Bwd(1)"[#HMI_No];
   "Control_DB".LCnv_Sys[#System_No].Cnv_Level[#Level].Cnv1.Instruction.Mode_Change := "CNV_HMI"."Mode_Change(1)"[#HMI_No];
   "Control_DB".LCnv_Sys[#System_No].Cnv_Level[#Level].Cnv1.Instruction.Enable := "CNV_HMI"."Enable(1)"[#HMI_No];
   #Light_Guard_Bypass := "HMI_Light_Guard_Bypass";

   "Control_DB".LCnv_Sys[#System_No].Cnv_Level[#Level].Cnv1.Instruction.Reset := "CNV_HMI"."Reset(1)"[#HMI_No] OR "Screen_DB_1".Reset_All[#HMI_No];
   IF "Control_DB".LCnv_Sys[#System_No].Cnv_Level[#Level].Cnv1.Mode <> 3 THEN
       "Control_DB".LCnv_Sys[#System_No].Cnv_Level[#Level].Cnv1.Instruction.Foward := "CNV_HMI"."Manual_Fwd(1)"[#HMI_No];
       "Control_DB".LCnv_Sys[#System_No].Cnv_Level[#Level].Cnv1.Instruction.Backward := "CNV_HMI"."Manual_Bwd(1)"[#HMI_No];
       "Control_DB".LCnv_Sys[#System_No].Cnv_Level[#Level].Cnv1.Instruction.Start_Transfer := "CNV_HMI"."Start_Transfer(1)"[#HMI_No];
       "Control_DB".LCnv_Sys[#System_No].Cnv_Level[#Level].Cnv1.Safety_Stop_Cnrl.Instruction.Manual_Extend := "CNV_HMI"."Manual_Sfty_Stopper_Up(1)"[#HMI_No];
       "Control_DB".LCnv_Sys[#System_No].Cnv_Level[#Level].Cnv1.Safety_Stop_Cnrl.Instruction.Manual_Retract := "CNV_HMI"."Manual_Sfty_Stopper_Down(1)"[#HMI_No];
       "Control_DB".LCnv_Sys[#System_No].Cnv_Level[#Level].Cnv1.Instruction.Task_ID := "CNV_HMI"."Task_ID(1)"[#HMI_No];
       "Control_DB".LCnv_Sys[#System_No].Cnv_Level[#Level].Cnv1.Instruction.Pallet_Align_Left := "CNV_HMI"."Pallet_Align_Left(1)"[#HMI_No];
       "Control_DB".LCnv_Sys[#System_No].Cnv_Level[#Level].Cnv1.Instruction.Pallet_Align_Right := "CNV_HMI"."Pallet_Align_Right(1)"[#HMI_No];
       IF "CNV_HMI"."Mode_Change(1)"[#HMI_No] <> 2 THEN
           "Control_DB".LCnv_Sys[#System_No].Cnv_Level[#Level].Cnv1.Instruction.Pallet_Allignment := "CNV_HMI"."Pallet_Allignment(1)"[#HMI_No] := FALSE;
       ELSE
           "Control_DB".LCnv_Sys[#System_No].Cnv_Level[#Level].Cnv1.Instruction.Pallet_Allignment := "CNV_HMI"."Pallet_Allignment(1)"[#HMI_No];
       END_IF;
       IF "CNV_HMI".In_Out[#HMI_No] THEN // 0 = ECNV RECEIVE, 1 = ECONV SEND
           "Control_DB".LCnv_Sys[#System_No].Cnv_Level[#Level].Cnv1.Instruction.Transfer_To_ID := 0;
           "Control_DB".LCnv_Sys[#System_No].Cnv_Level[#Level].Cnv1.Instruction.Transfer_From_ID := DINT#120000 + (#Level * 100) + #System_No;
       ELSE
           "Control_DB".LCnv_Sys[#System_No].Cnv_Level[#Level].Cnv1.Instruction.Transfer_To_ID := DINT#120000 + (#Level * 100) + #System_No;
           "Control_DB".LCnv_Sys[#System_No].Cnv_Level[#Level].Cnv1.Instruction.Transfer_From_ID := 0;
       END_IF;
   END_IF;
END_FUNCTION

FUNCTION "Feed_BCNV_Cnv1" : Void   // FC31, SCL
{ S7_Optimized_Access := 'TRUE' }
VERSION : 0.1
// stored: AutoNumber true, IsIECCheckEnabled false, SetENOAutomatically false, UDAEnableTagReadback false
   VAR_INPUT
      System_No : UInt;
      Level : UInt;
   END_VAR
BEGIN
   //Sensors
   "HMI_CNV_Left" := "Control_DB".LCnv_Sys[#System_No].Cnv_Level[#Level].Cnv1.Inputs.Left;
   "HMI_CNV_Lpd1" := "Control_DB".LCnv_Sys[#System_No].Cnv_Level[#Level].Cnv1.Inputs.Lpd1;
   "HMI_CNV_Lpd2" := "Control_DB".LCnv_Sys[#System_No].Cnv_Level[#Level].Cnv1.Inputs.Lpd2;
   "HMI_CNV_Right" := "Control_DB".LCnv_Sys[#System_No].Cnv_Level[#Level].Cnv1.Inputs.Right;
   "HMI_CNV_Rpd1" := "Control_DB".LCnv_Sys[#System_No].Cnv_Level[#Level].Cnv1.Inputs.Rpd1;
   "HMI_CNV_Rpd2" := "Control_DB".LCnv_Sys[#System_No].Cnv_Level[#Level].Cnv1.Inputs.Rpd2;"HMI_CNV_Sdetect1" := "Control_DB".LCnv_Sys[#System_No].Cnv_Level[#Level].Cnv1.Inputs.Sdetect1;
   "HMI_CNV_Sdetect2" := "Control_DB".LCnv_Sys[#System_No].Cnv_Level[#Level].Cnv1.Inputs.Sdetect2;
   "HMI_CNV_SftyPinUp" := "Control_DB".LCnv_Sys[#System_No].Cnv_Level[#Level].Cnv1.Safety_Stop_Cnrl.Inputs.DP_Extended;
   "HMI_CNV_SftyPinDown" := "Control_DB".LCnv_Sys[#System_No].Cnv_Level[#Level].Cnv1.Safety_Stop_Cnrl.Inputs.DP_Retracted;
   IF "Control_DB".LCnv_Sys[#System_No].Cnv_Level[#Level].Cnv1.Safety_Stop_Cnrl.Inputs.DP_Extended AND
       NOT "Control_DB".LCnv_Sys[#System_No].Cnv_Level[#Level].Cnv1.Safety_Stop_Cnrl.Inputs.DP_Retracted THEN
       "UpDown" := 1;
   ELSIF NOT "Control_DB".LCnv_Sys[#System_No].Cnv_Level[#Level].Cnv1.Safety_Stop_Cnrl.Inputs.DP_Extended AND
       "Control_DB".LCnv_Sys[#System_No].Cnv_Level[#Level].Cnv1.Safety_Stop_Cnrl.Inputs.DP_Retracted THEN
       "UpDown" := 2;
   ELSE
       "UpDown" := 0;
   END_IF;

   //Feedback
   "Mode_HMI" := "Control_DB".LCnv_Sys[#System_No].Cnv_Level[#Level].Cnv1.Mode;
   "Enabled_HMI" := "Control_DB".LCnv_Sys[#System_No].Cnv_Level[#Level].Cnv1.Enabled;
   "Error_HMI" := "Control_DB".LCnv_Sys[#System_No].Cnv_Level[#Level].Cnv1.Error;
   "Warning_HMI" := "Control_DB".LCnv_Sys[#System_No].Cnv_Level[#Level].Cnv1.Warning;
   "Stopped_HMI" := "Control_DB".LCnv_Sys[#System_No].Cnv_Level[#Level].Cnv1.Stopped;
   "Running_HMI" := "Control_DB".LCnv_Sys[#System_No].Cnv_Level[#Level].Cnv1.Running;
   "Ready_For_Task_HMI" := "Control_DB".LCnv_Sys[#System_No].Cnv_Level[#Level].Cnv1.Ready_For_Task;
   "Cnv_Occupied_HMI" := "Control_DB".LCnv_Sys[#System_No].Cnv_Level[#Level].Cnv1.Cnv_Occupied;
   "Shuttle_in_place_HMI" := "Control_DB".LCnv_Sys[#System_No].Cnv_Level[#Level].Cnv1.Shuttle_In_Place;
   "Current_Task_Type_HMI" := "Control_DB".LCnv_Sys[#System_No].Cnv_Level[#Level].Cnv1.Current_Task_Type;
   "Current_Task_ID_HMI" := "Control_DB".LCnv_Sys[#System_No].Cnv_Level[#Level].Cnv1.Current_Task_ID;
   "SM_State_HMI" := "Control_DB".LCnv_Sys[#System_No].Cnv_Level[#Level].Cnv1.SM_State;
   IF "Control_DB".LCnv_Sys[#System_No].Cnv_Level[#Level].Cnv1.Motor.Forward THEN
       "Motor_Direction_HMI" := 1;
   ELSIF "Control_DB".LCnv_Sys[#System_No].Cnv_Level[#Level].Cnv1.Motor.Reverse THEN
       "Motor_Direction_HMI" := 2;
   ELSE
       "Motor_Direction_HMI" := 0;
   END_IF;
   "Motor_Speed_Requested_HMI" := "Control_DB".LCnv_Sys[#System_No].Cnv_Level[#Level].Cnv1.Motor.Speed;
   "Motor_Speed_Actual_HMI" := "Control_DB".LCnv_Sys[#System_No].Cnv_Level[#Level].Cnv1.Motor.Speed_Actual;
   "Transfer_To_ID_HMI" := "Control_DB".LCnv_Sys[#System_No].Cnv_Level[#Level].Cnv1.Instruction.Transfer_To_ID;
   "Transfer_From_ID_HMI" := "Control_DB".LCnv_Sys[#System_No].Cnv_Level[#Level].Cnv1.Instruction.Transfer_From_ID;

   //Instructions
   "Control_DB".LCnv_Sys[#System_No].Cnv_Level[#Level].Cnv1.Instruction.Stop := "Stop_HMI";
   "Control_DB".LCnv_Sys[#System_No].Cnv_Level[#Level].Cnv1.Instruction.Execute := "Manual_Fwd_HMI" OR "Manual_Bwd_HMI";
   "Control_DB".LCnv_Sys[#System_No].Cnv_Level[#Level].Cnv1.Instruction.Mode_Change := "Mode_Change_HMI";
   "Control_DB".LCnv_Sys[#System_No].Cnv_Level[#Level].Cnv1.Instruction.Enable := "Enable_HMI";
   "Control_DB".LCnv_Sys[#System_No].Cnv_Level[#Level].Cnv1.Instruction.Reset := "Reset_HMI";
   IF "Control_DB".LCnv_Sys[#System_No].Cnv_Level[#Level].Cnv1.Mode <> 3 THEN
       "Control_DB".LCnv_Sys[#System_No].Cnv_Level[#Level].Cnv1.Instruction.Foward := "Manual_Fwd_HMI";
       "Control_DB".LCnv_Sys[#System_No].Cnv_Level[#Level].Cnv1.Instruction.Backward := "Manual_Bwd_HMI";
       "Control_DB".LCnv_Sys[#System_No].Cnv_Level[#Level].Cnv1.Instruction.Start_Transfer := "Start_Transfer_HMI";
       IF "Control_DB".LCnv_Sys[#System_No].Cnv_Level[#Level].Cnv1.Mode = 1 THEN
           "Control_DB".LCnv_Sys[#System_No].Cnv_Level[#Level].Cnv1.Instruction.Start_Transfer_Backward := "Transfer_Backward";
       END_IF;
       "Control_DB".LCnv_Sys[#System_No].Cnv_Level[#Level].Cnv1.Safety_Stop_Cnrl.Instruction.Manual_Extend := "Manual_Sfty_Stopper_Up";
       "Control_DB".LCnv_Sys[#System_No].Cnv_Level[#Level].Cnv1.Safety_Stop_Cnrl.Instruction.Manual_Retract := "Manual_Sfty_Stopper_Down";
       "Control_DB".LCnv_Sys[#System_No].Cnv_Level[#Level].Cnv1.Instruction.Task_ID := "Task_ID_HMI";
       "Control_DB".LCnv_Sys[#System_No].Cnv_Level[#Level].Cnv1.Instruction.Pallet_Align_Left := "Pallet_Align_Left_HMI";
       "Control_DB".LCnv_Sys[#System_No].Cnv_Level[#Level].Cnv1.Instruction.Pallet_Align_Right := "Pallet_Align_Right_HMI";
       "Control_DB".LCnv_Sys[#System_No].Cnv_Level[#Level].Cnv1.Instruction.Pallet_Allignment := "Pallet_Align_Right_HMI";
       IF "CNV_HMI".In_Out[#System_No] THEN // 0 = Inbound, 1 = Outbound
           "Control_DB".LCnv_Sys[#System_No].Cnv_Level[#Level].Cnv1.Instruction.Transfer_To_ID := DINT#100000 + (#Level * 100) + #System_No;
           "Control_DB".LCnv_Sys[#System_No].Cnv_Level[#Level].Cnv1.Instruction.Transfer_From_ID := 0;
       ELSE
           "Control_DB".LCnv_Sys[#System_No].Cnv_Level[#Level].Cnv1.Instruction.Transfer_To_ID := 0;
           "Control_DB".LCnv_Sys[#System_No].Cnv_Level[#Level].Cnv1.Instruction.Transfer_From_ID := DINT#100000 + (#Level * 100+ #System_No);
       END_IF;
   END_IF;
END_FUNCTION

FUNCTION "Feed_BCNV_Cnv2(1)" : Void   // FC28, SCL
{ S7_Optimized_Access := 'TRUE' }
VERSION : 0.1
// stored: AutoNumber true, IsIECCheckEnabled false, SetENOAutomatically false, UDAEnableTagReadback false
   VAR_INPUT
      System_No : UInt;
      Level : UInt;
      Light_Guard_IO : Bool;
   END_VAR
   VAR_OUTPUT
      Light_Guard_Bypass : Bool;
   END_VAR
   VAR_IN_OUT
      System_Busy : Bool;
   END_VAR
BEGIN
   //Sensors
   "HMI_CNV_Left(1)" := "Control_DB".LCnv_Sys[#System_No].Cnv_Level[#Level].Cnv2.Inputs.Left;
   "HMI_CNV_Lpd1(1)" := "Control_DB".LCnv_Sys[#System_No].Cnv_Level[#Level].Cnv2.Inputs.Lpd1;
   "HMI_CNV_Lpd2(1)" := "Control_DB".LCnv_Sys[#System_No].Cnv_Level[#Level].Cnv2.Inputs.Lpd2;
   "HMI_CNV_Right(1)" := "Control_DB".LCnv_Sys[#System_No].Cnv_Level[#Level].Cnv2.Inputs.Right;
   "HMI_CNV_Rpd1(1)" := "Control_DB".LCnv_Sys[#System_No].Cnv_Level[#Level].Cnv2.Inputs.Rpd1;
   "HMI_CNV_Rpd2(1)" := "Control_DB".LCnv_Sys[#System_No].Cnv_Level[#Level].Cnv2.Inputs.Rpd2;
   "HMI_CNV_Sdetect1(1)" := "Control_DB".LCnv_Sys[#System_No].Cnv_Level[#Level].Cnv2.Inputs.Sdetect1;
   "HMI_CNV_Sdetect2(1)" := "Control_DB".LCnv_Sys[#System_No].Cnv_Level[#Level].Cnv2.Inputs.Sdetect2;
   "HMI_CNV_SftyPinUp(1)" := "Control_DB".LCnv_Sys[#System_No].Cnv_Level[#Level].Cnv2.Safety_Stop_Cnrl.Inputs.DP_Extended;
   "HMI_CNV_SftyPinDown(1)" := "Control_DB".LCnv_Sys[#System_No].Cnv_Level[#Level].Cnv2.Safety_Stop_Cnrl.Inputs.DP_Retracted;
   "HMI_Light_Guard" := #System_No <= 3 AND #Level = 1 AND "HMI_DB".Username = 'admin'; //To show the button
   IF "Control_DB".LCnv_Sys[#System_No].Cnv_Level[#Level].Cnv2.Safety_Stop_Cnrl.Inputs.DP_Extended AND
       NOT "Control_DB".LCnv_Sys[#System_No].Cnv_Level[#Level].Cnv2.Safety_Stop_Cnrl.Inputs.DP_Retracted THEN
       "UpDown(1)" := 1;
   ELSIF NOT "Control_DB".LCnv_Sys[#System_No].Cnv_Level[#Level].Cnv2.Safety_Stop_Cnrl.Inputs.DP_Extended AND
       "Control_DB".LCnv_Sys[#System_No].Cnv_Level[#Level].Cnv2.Safety_Stop_Cnrl.Inputs.DP_Retracted THEN
       "UpDown(1)" := 2;
   ELSE
       "UpDown(1)" := 0;
   END_IF;

   //Status
   "Mode_HMI(1)" := "Control_DB".LCnv_Sys[#System_No].Cnv_Level[#Level].Cnv2.Mode;
   "Enabled_HMI(1)" := "Control_DB".LCnv_Sys[#System_No].Cnv_Level[#Level].Cnv2.Enabled;
   "Error_HMI(1)" := "Control_DB".LCnv_Sys[#System_No].Cnv_Level[#Level].Cnv2.Error;
   "Warning_HMI(1)" := "Control_DB".LCnv_Sys[#System_No].Cnv_Level[#Level].Cnv2.Warning;
   "Stopped_HMI(1)" := "Control_DB".LCnv_Sys[#System_No].Cnv_Level[#Level].Cnv2.Stopped;
   "Running_HMI(1)" := "Control_DB".LCnv_Sys[#System_No].Cnv_Level[#Level].Cnv2.Running;
   "Ready_For_Task_HMI(1)" := "Control_DB".LCnv_Sys[#System_No].Cnv_Level[#Level].Cnv2.Ready_For_Task;
   "Cnv_Occupied_HMI(1)" := "Control_DB".LCnv_Sys[#System_No].Cnv_Level[#Level].Cnv2.Cnv_Occupied;
   "Shuttle_in_place_HMI(1)" := "Control_DB".LCnv_Sys[#System_No].Cnv_Level[#Level].Cnv2.Shuttle_In_Place;
   "Current_Task_Type_HMI(1)" := "Control_DB".LCnv_Sys[#System_No].Cnv_Level[#Level].Cnv2.Current_Task_Type;
   "Current_Task_ID_HMI(1)" := "Control_DB".LCnv_Sys[#System_No].Cnv_Level[#Level].Cnv2.Current_Task_ID;
   "SM_State_HMI(1)" := "Control_DB".LCnv_Sys[#System_No].Cnv_Level[#Level].Cnv2.SM_State;
   "Pallet_Type_HMI(1)" := "Control_DB".LCnv_Sys[#System_No].Cnv_Level[#Level].Cnv2.Pallet_Type;
   IF "Control_DB".LCnv_Sys[#System_No].Cnv_Level[#Level].Cnv2.Motor.Forward THEN
       "Motor_Direction_HMI(1)" := 1;
   ELSIF "Control_DB".LCnv_Sys[#System_No].Cnv_Level[#Level].Cnv2.Motor.Reverse THEN
       "Motor_Direction_HMI(1)" := 2;
   ELSE
       "Motor_Direction_HMI(1)" := 0;
   END_IF;
   "Motor_Speed_Requested_HMI(1)" := "Control_DB".LCnv_Sys[#System_No].Cnv_Level[#Level].Cnv2.Motor.Speed;
   "Motor_Speed_Actual_HMI(1)" := "Control_DB".LCnv_Sys[#System_No].Cnv_Level[#Level].Cnv2.Motor.Speed_Actual;
   "CNV_Motor_Ready(1)" := "Control_DB".LCnv_Sys[#System_No].Cnv_Level[#Level].Cnv2.Motor.Ready;
   "CNV_Motor_Current_Actual_HMI(1)" := "Control_DB".LCnv_Sys[#System_No].Cnv_Level[#Level].Cnv2.Motor.Actual_Current;
   "CNV_Motor_Actual_Torque(1)" := "Control_DB".LCnv_Sys[#System_No].Cnv_Level[#Level].Cnv2.Motor.Actual_Torque;
   "Transfer_To_ID_HMI(1)" := "Control_DB".LCnv_Sys[#System_No].Cnv_Level[#Level].Cnv2.Instruction.Transfer_To_ID;
   "Transfer_From_ID_HMI(1)" := "Control_DB".LCnv_Sys[#System_No].Cnv_Level[#Level].Cnv2.Instruction.Transfer_From_ID;

   IF "Control_DB".LCnv_Sys[#System_No].Cnv_Level[#Level].Cnv2.Motor.Error THEN
       "CNV_Motor_Status_HMI(1)" := 2;
   ELSIF "Control_DB".LCnv_Sys[#System_No].Cnv_Level[#Level].Cnv2.Motor.Enabled THEN
       "CNV_Motor_Status_HMI(1)" := 1;
   ELSIF NOT "Control_DB".LCnv_Sys[#System_No].Cnv_Level[#Level].Cnv2.Motor.Enabled THEN
       "CNV_Motor_Status_HMI(1)" := 0;
   END_IF;

   //Instructions
   IF ("HMI_Box_Connected_1" = #System_No OR ("HMI_Box_Connected_1" >= (#System_No * 10) + 1 AND "HMI_Box_Connected_1" <= (#System_No * 10) + 8)) OR
       ("HMI_Box_Connected_2" = #System_No OR ("HMI_Box_Connected_1" >= (#System_No * 10) + 1 AND "HMI_Box_Connected_1" <= (#System_No * 10) + 8))
   THEN
       #System_Busy := TRUE;
   ELSE
       #System_Busy := FALSE;
       "Control_DB".LCnv_Sys[#System_No].Cnv_Level[#Level].Cnv2.Instruction.Stop := "Stop_HMI(1)";
       "Control_DB".LCnv_Sys[#System_No].Cnv_Level[#Level].Cnv2.Instruction.Execute := "Manual_Fwd_HMI(1)" OR "Manual_Bwd_HMI(1)";
       IF "BT_Confirmation_HMI" THEN
           "Control_DB".VTD_Sys[#System_No].Instruction.Mode_Change :=
           "Control_DB".ECnv_Sys[#System_No].Instruction.Mode_Change :=
           "Control_DB".LCnv_Sys[#System_No].Cnv_Level[1].Cnv1.Instruction.Mode_Change :=
           "Control_DB".LCnv_Sys[#System_No].Cnv_Level[2].Cnv1.Instruction.Mode_Change :=
           "Control_DB".LCnv_Sys[#System_No].Cnv_Level[3].Cnv1.Instruction.Mode_Change :=
           "Control_DB".LCnv_Sys[#System_No].Cnv_Level[4].Cnv1.Instruction.Mode_Change :=
           "Control_DB".LCnv_Sys[#System_No].Cnv_Level[5].Cnv1.Instruction.Mode_Change :=
           "Control_DB".LCnv_Sys[#System_No].Cnv_Level[6].Cnv1.Instruction.Mode_Change :=
           "Control_DB".LCnv_Sys[#System_No].Cnv_Level[7].Cnv1.Instruction.Mode_Change :=
           "Control_DB".LCnv_Sys[#System_No].Cnv_Level[8].Cnv1.Instruction.Mode_Change :=
           "Control_DB".LCnv_Sys[#System_No].Cnv_Level[1].Cnv2.Instruction.Mode_Change :=
           "Control_DB".LCnv_Sys[#System_No].Cnv_Level[2].Cnv2.Instruction.Mode_Change :=
           "Control_DB".LCnv_Sys[#System_No].Cnv_Level[3].Cnv2.Instruction.Mode_Change :=
           "Control_DB".LCnv_Sys[#System_No].Cnv_Level[4].Cnv2.Instruction.Mode_Change :=
           "Control_DB".LCnv_Sys[#System_No].Cnv_Level[5].Cnv2.Instruction.Mode_Change :=
           "Control_DB".LCnv_Sys[#System_No].Cnv_Level[6].Cnv2.Instruction.Mode_Change :=
           "Control_DB".LCnv_Sys[#System_No].Cnv_Level[7].Cnv2.Instruction.Mode_Change :=
           "Control_DB".LCnv_Sys[#System_No].Cnv_Level[8].Cnv2.Instruction.Mode_Change := "Mode_Change_HMI(1)";
           "Mode_Change_HMI" := "Mode_Change_HMI(1)";
           "BT_Confirmation_HMI" := FALSE;
       END_IF;

       "Control_DB".LCnv_Sys[#System_No].Cnv_Level[#Level].Cnv2.Instruction.Enable := "Enable_HMI(1)";
       IF "Control_DB".LCnv_Sys[#System_No].Cnv_Level[#Level].Cnv1.Mode <> 1 THEN
           "HMI_Light_Guard_Bypass" := FALSE;
       ELSIF "HMI_Light_Guard_Bypass" AND "Control_DB".LCnv_Sys[#System_No].Cnv_Level[1].Cnv1.Error THEN
           #Light_Guard_Bypass := TRUE;
       ELSIF NOT "Control_DB".LCnv_Sys[#System_No].Cnv_Level[1].Cnv1.Running AND NOT "Control_DB".LCnv_Sys[#System_No].Cnv_Level[1].Cnv1.Error AND #Light_Guard_IO THEN //Not Running and No error and light guard free
           #Light_Guard_Bypass := FALSE; //Cancel bypass
       END_IF;

       "Control_DB".LCnv_Sys[#System_No].Cnv_Level[#Level].Cnv2.Instruction.Reset :=
       "Reset_HMI(1)" OR "Reset_All" OR
       "CNV_HMI"."Reset(1)"[1] OR "Screen_DB_1".Reset_All[1] OR
       "CNV_HMI"."Reset(1)"[2] OR "Screen_DB_1".Reset_All[2];

       IF "Control_DB".LCnv_Sys[#System_No].Cnv_Level[#Level].Cnv2.Mode <> 3 THEN
           "Control_DB".LCnv_Sys[#System_No].Cnv_Level[#Level].Cnv2.Instruction.Foward := "Manual_Fwd_HMI(1)";
           "Control_DB".LCnv_Sys[#System_No].Cnv_Level[#Level].Cnv2.Instruction.Backward := "Manual_Bwd_HMI(1)";
           "Control_DB".LCnv_Sys[#System_No].Cnv_Level[#Level].Cnv2.Instruction.Start_Transfer := "Start_Transfer_HMI(1)";
           IF "Control_DB".LCnv_Sys[#System_No].Cnv_Level[#Level].Cnv2.Mode = 1 THEN
               "Control_DB".LCnv_Sys[#System_No].Cnv_Level[#Level].Cnv2.Instruction.Start_Transfer_Backward := "Transfer_Backward(1)";
           END_IF;
           "Control_DB".LCnv_Sys[#System_No].Cnv_Level[#Level].Cnv2.Safety_Stop_Cnrl.Instruction.Manual_Extend := "Manual_Sfty_Stopper_Up(1)";
           "Control_DB".LCnv_Sys[#System_No].Cnv_Level[#Level].Cnv2.Safety_Stop_Cnrl.Instruction.Manual_Retract := "Manual_Sfty_Stopper_Down(1)";
           "Control_DB".LCnv_Sys[#System_No].Cnv_Level[#Level].Cnv2.Instruction.Task_ID := "Task_ID_HMI(1)";
           "Control_DB".LCnv_Sys[#System_No].Cnv_Level[#Level].Cnv2.Instruction.Pallet_Align_Left := "Pallet_Align_Left_HMI(1)";
           "Control_DB".LCnv_Sys[#System_No].Cnv_Level[#Level].Cnv2.Instruction.Pallet_Align_Right := "Pallet_Align_Right_HMI(1)";
           IF "Mode_Change_HMI(1)" <> 2 THEN
               "Control_DB".LCnv_Sys[#System_No].Cnv_Level[#Level].Cnv2.Instruction.Pallet_Allignment := "Pallet_Allignment_HMI(1)" := FALSE;
           ELSE
               "Control_DB".LCnv_Sys[#System_No].Cnv_Level[#Level].Cnv2.Instruction.Pallet_Allignment := "Pallet_Allignment_HMI(1)";
           END_IF;
           IF "CNV_HMI".In_Out[#System_No] THEN // 0 = ECNV RECEIVE, 1 = ECONV SEND
               "Control_DB".LCnv_Sys[#System_No].Cnv_Level[#Level].Cnv2.Instruction.Transfer_To_ID := 0;
               "Control_DB".LCnv_Sys[#System_No].Cnv_Level[#Level].Cnv2.Instruction.Transfer_From_ID := DINT#120000 + (#Level * 100) + #System_No;
           ELSE
               "Control_DB".LCnv_Sys[#System_No].Cnv_Level[#Level].Cnv2.Instruction.Transfer_To_ID := DINT#120000 + (#Level * 100) + #System_No;
               "Control_DB".LCnv_Sys[#System_No].Cnv_Level[#Level].Cnv2.Instruction.Transfer_From_ID := 0;
           END_IF;
       END_IF;
   END_IF;
END_FUNCTION

FUNCTION "Feed_BCNV_Cnv2(1)_1" : Void   // FC30, SCL
{ S7_Optimized_Access := 'TRUE' }
VERSION : 0.1
// stored: AutoNumber true, IsIECCheckEnabled false, SetENOAutomatically false, UDAEnableTagReadback false
   VAR_INPUT
      HMI_No : UInt;
      System_No : UInt;
      Level : UInt;
      Light_Guard_IO : Bool;
   END_VAR
   VAR_OUTPUT
      Light_Guard_Bypass : Bool;
   END_VAR
BEGIN
   //Sensors
   "CNV_HMI"."Left(1)"[#HMI_No] := "Control_DB".LCnv_Sys[#System_No].Cnv_Level[#Level].Cnv2.Inputs.Left;
   "CNV_HMI"."Lpd1(1)"[#HMI_No] := "Control_DB".LCnv_Sys[#System_No].Cnv_Level[#Level].Cnv2.Inputs.Lpd1;
   "CNV_HMI"."Lpd2(1)"[#HMI_No] := "Control_DB".LCnv_Sys[#System_No].Cnv_Level[#Level].Cnv2.Inputs.Lpd2;
   "CNV_HMI"."Right(1)"[#HMI_No] := "Control_DB".LCnv_Sys[#System_No].Cnv_Level[#Level].Cnv2.Inputs.Right;
   "CNV_HMI"."Rpd1(1)"[#HMI_No] := "Control_DB".LCnv_Sys[#System_No].Cnv_Level[#Level].Cnv2.Inputs.Rpd1;
   "CNV_HMI"."Rpd2(1)"[#HMI_No] := "Control_DB".LCnv_Sys[#System_No].Cnv_Level[#Level].Cnv2.Inputs.Rpd2;
   "CNV_HMI"."Sdetect1(1)"[#HMI_No] := "Control_DB".LCnv_Sys[#System_No].Cnv_Level[#Level].Cnv2.Inputs.Sdetect1;
   "CNV_HMI"."Sdetect2(1)"[#HMI_No] := "Control_DB".LCnv_Sys[#System_No].Cnv_Level[#Level].Cnv2.Inputs.Sdetect2;
   "HMI_Light_Guard" := #Level = 1; //To show the button
   IF "Control_DB".LCnv_Sys[#System_No].Cnv_Level[#Level].Cnv2.Safety_Stop_Cnrl.Inputs.DP_Extended AND
       NOT "Control_DB".LCnv_Sys[#System_No].Cnv_Level[#Level].Cnv2.Safety_Stop_Cnrl.Inputs.DP_Retracted THEN
       "CNV_HMI"."UpDown(1)"[#HMI_No] := 1;
   ELSIF NOT "Control_DB".LCnv_Sys[#System_No].Cnv_Level[#Level].Cnv2.Safety_Stop_Cnrl.Inputs.DP_Extended AND
       "Control_DB".LCnv_Sys[#System_No].Cnv_Level[#Level].Cnv2.Safety_Stop_Cnrl.Inputs.DP_Retracted THEN
       "CNV_HMI"."UpDown(1)"[#HMI_No] := 2;
   ELSE
       "CNV_HMI"."UpDown(1)"[#HMI_No] := 0;
   END_IF;

   //Status
   "CNV_HMI"."Mode(1)"[#HMI_No] := "Control_DB".LCnv_Sys[#System_No].Cnv_Level[#Level].Cnv2.Mode;
   "CNV_HMI"."Enabled(1)"[#HMI_No] := "Control_DB".LCnv_Sys[#System_No].Cnv_Level[#Level].Cnv2.Enabled;
   "CNV_HMI"."Error(1)"[#HMI_No] := "Control_DB".LCnv_Sys[#System_No].Cnv_Level[#Level].Cnv2.Error;
   "CNV_HMI"."Warning(1)"[#HMI_No] := "Control_DB".LCnv_Sys[#System_No].Cnv_Level[#Level].Cnv2.Warning;
   "CNV_HMI"."Stopped(1)"[#HMI_No] := "Control_DB".LCnv_Sys[#System_No].Cnv_Level[#Level].Cnv2.Stopped;
   "CNV_HMI"."Running(1)"[#HMI_No] := "Control_DB".LCnv_Sys[#System_No].Cnv_Level[#Level].Cnv2.Running;
   "CNV_HMI"."Ready_For_Task(1)"[#HMI_No] := "Control_DB".LCnv_Sys[#System_No].Cnv_Level[#Level].Cnv2.Ready_For_Task;
   "CNV_HMI"."Occupied(1)"[#HMI_No] := "Control_DB".LCnv_Sys[#System_No].Cnv_Level[#Level].Cnv2.Cnv_Occupied;
   "CNV_HMI"."Shuttle_in_place(1)"[#HMI_No] := "Control_DB".LCnv_Sys[#System_No].Cnv_Level[#Level].Cnv2.Shuttle_In_Place;
   "CNV_HMI"."Current_Task_Type(1)"[#HMI_No] := "Control_DB".LCnv_Sys[#System_No].Cnv_Level[#Level].Cnv2.Current_Task_Type;
   "CNV_HMI"."Task_ID(1)"[#HMI_No] := "Control_DB".LCnv_Sys[#System_No].Cnv_Level[#Level].Cnv2.Current_Task_ID;
   "CNV_HMI"."SM_State(1)"[#HMI_No] := "Control_DB".LCnv_Sys[#System_No].Cnv_Level[#Level].Cnv2.SM_State;
   "CNV_HMI"."Pallet_Type(1)"[#HMI_No] := "Control_DB".LCnv_Sys[#System_No].Cnv_Level[#Level].Cnv2.Pallet_Type;
   IF "Control_DB".LCnv_Sys[#System_No].Cnv_Level[#Level].Cnv2.Motor.Forward THEN
       "CNV_HMI"."Motor_Direction(1)"[#HMI_No] := 1;
   ELSIF "Control_DB".LCnv_Sys[#System_No].Cnv_Level[#Level].Cnv2.Motor.Reverse THEN
       "CNV_HMI"."Motor_Direction(1)"[#HMI_No] := 2;
   ELSE
       "CNV_HMI"."Motor_Direction(1)"[#HMI_No] := 0;
   END_IF;
   "CNV_HMI"."Motor_Speed_Requested(1)"[#HMI_No] := "Control_DB".LCnv_Sys[#System_No].Cnv_Level[#Level].Cnv2.Motor.Speed;
   "CNV_HMI"."Motor_Speed_Actual(1)"[#HMI_No] := "Control_DB".LCnv_Sys[#System_No].Cnv_Level[#Level].Cnv2.Motor.Speed_Actual;
   "CNV_HMI"."Motor_Ready(1)"[#HMI_No] := "Control_DB".LCnv_Sys[#System_No].Cnv_Level[#Level].Cnv2.Motor.Ready;
   "CNV_HMI"."Motor_Current_Actual(1)"[#HMI_No] := "Control_DB".LCnv_Sys[#System_No].Cnv_Level[#Level].Cnv2.Motor.Actual_Current;
   "CNV_HMI"."Motor_Actual_Torque(1)"[#HMI_No] := "Control_DB".LCnv_Sys[#System_No].Cnv_Level[#Level].Cnv2.Motor.Actual_Torque;
   "CNV_HMI"."Transfer_To_ID(1)"[#HMI_No] := "Control_DB".LCnv_Sys[#System_No].Cnv_Level[#Level].Cnv2.Instruction.Transfer_To_ID;
   "CNV_HMI"."Transfer_From_ID(1)"[#HMI_No] := "Control_DB".LCnv_Sys[#System_No].Cnv_Level[#Level].Cnv2.Instruction.Transfer_From_ID;

   IF "Control_DB".LCnv_Sys[#System_No].Cnv_Level[#Level].Cnv2.Motor.Error THEN
       "CNV_HMI"."Motor_Status(1)"[#HMI_No] := 2;
   ELSIF "Control_DB".LCnv_Sys[#System_No].Cnv_Level[#Level].Cnv2.Motor.Enabled THEN
       "CNV_HMI"."Motor_Status(1)"[#HMI_No] := 1;
   ELSIF NOT "Control_DB".LCnv_Sys[#System_No].Cnv_Level[#Level].Cnv2.Motor.Enabled THEN
       "CNV_HMI"."Motor_Status(1)"[#HMI_No] := 0;
   END_IF;

   //Instructions
   "Control_DB".LCnv_Sys[#System_No].Cnv_Level[#Level].Cnv2.Instruction.Stop := "CNV_HMI"."Stop(1)"[#HMI_No];
   "Control_DB".LCnv_Sys[#System_No].Cnv_Level[#Level].Cnv2.Instruction.Execute := "CNV_HMI"."Manual_Fwd(1)"[#HMI_No] OR "CNV_HMI"."Manual_Bwd(1)"[#HMI_No];
   "Control_DB".LCnv_Sys[#System_No].Cnv_Level[#Level].Cnv2.Instruction.Mode_Change := "CNV_HMI"."Mode_Change(1)"[#HMI_No];
   "Control_DB".LCnv_Sys[#System_No].Cnv_Level[#Level].Cnv2.Instruction.Enable := "CNV_HMI"."Enable(1)"[#HMI_No];
   #Light_Guard_Bypass := "HMI_Light_Guard_Bypass";

   "Control_DB".LCnv_Sys[#System_No].Cnv_Level[#Level].Cnv2.Instruction.Reset := "CNV_HMI"."Reset(1)"[#HMI_No] OR "Screen_DB_1".Reset_All[#HMI_No];
   IF "Control_DB".LCnv_Sys[#System_No].Cnv_Level[#Level].Cnv2.Mode <> 3 THEN
       "Control_DB".LCnv_Sys[#System_No].Cnv_Level[#Level].Cnv2.Instruction.Foward := "CNV_HMI"."Manual_Fwd(1)"[#HMI_No];
       "Control_DB".LCnv_Sys[#System_No].Cnv_Level[#Level].Cnv2.Instruction.Backward := "CNV_HMI"."Manual_Bwd(1)"[#HMI_No];
       "Control_DB".LCnv_Sys[#System_No].Cnv_Level[#Level].Cnv2.Instruction.Start_Transfer := "CNV_HMI"."Start_Transfer(1)"[#HMI_No];
       "Control_DB".LCnv_Sys[#System_No].Cnv_Level[#Level].Cnv2.Safety_Stop_Cnrl.Instruction.Manual_Extend := "CNV_HMI"."Manual_Sfty_Stopper_Up(1)"[#HMI_No];
       "Control_DB".LCnv_Sys[#System_No].Cnv_Level[#Level].Cnv2.Safety_Stop_Cnrl.Instruction.Manual_Retract := "CNV_HMI"."Manual_Sfty_Stopper_Down(1)"[#HMI_No];
       "Control_DB".LCnv_Sys[#System_No].Cnv_Level[#Level].Cnv2.Instruction.Task_ID := "CNV_HMI"."Task_ID(1)"[#HMI_No];
       "Control_DB".LCnv_Sys[#System_No].Cnv_Level[#Level].Cnv2.Instruction.Pallet_Align_Left := "CNV_HMI"."Pallet_Align_Left(1)"[#HMI_No];
       "Control_DB".LCnv_Sys[#System_No].Cnv_Level[#Level].Cnv2.Instruction.Pallet_Align_Right := "CNV_HMI"."Pallet_Align_Right(1)"[#HMI_No];
       IF "CNV_HMI"."Mode_Change(1)"[#HMI_No] <> 2 THEN
           "Control_DB".LCnv_Sys[#System_No].Cnv_Level[#Level].Cnv2.Instruction.Pallet_Allignment := "CNV_HMI"."Pallet_Allignment(1)"[#HMI_No] := FALSE;
       ELSE
           "Control_DB".LCnv_Sys[#System_No].Cnv_Level[#Level].Cnv2.Instruction.Pallet_Allignment := "CNV_HMI"."Pallet_Allignment(1)"[#HMI_No];
       END_IF;
       IF "CNV_HMI".In_Out[#System_No] THEN // 0 = ECNV RECEIVE, 1 = ECONV SEND
           "Control_DB".LCnv_Sys[#System_No].Cnv_Level[#Level].Cnv2.Instruction.Transfer_To_ID := 0;
           "Control_DB".LCnv_Sys[#System_No].Cnv_Level[#Level].Cnv2.Instruction.Transfer_From_ID := DINT#120000 + (#Level * 100) + #System_No;
       ELSE
           "Control_DB".LCnv_Sys[#System_No].Cnv_Level[#Level].Cnv2.Instruction.Transfer_To_ID := DINT#120000 + (#Level * 100) + #System_No;
           "Control_DB".LCnv_Sys[#System_No].Cnv_Level[#Level].Cnv2.Instruction.Transfer_From_ID := 0;
       END_IF;
   END_IF;
END_FUNCTION

FUNCTION "Feed_BCNV_Cnv2" : Void   // FC32, SCL
{ S7_Optimized_Access := 'TRUE' }
VERSION : 0.1
// stored: AutoNumber true, IsIECCheckEnabled false, SetENOAutomatically false, UDAEnableTagReadback false
   VAR_INPUT
      System_No : UInt;
      Level : UInt;
   END_VAR
BEGIN
   //Sensors
   "HMI_CNV_Left" := "Control_DB".LCnv_Sys[#System_No].Cnv_Level[#Level].Cnv2.Inputs.Left;
   "HMI_CNV_Lpd1" := "Control_DB".LCnv_Sys[#System_No].Cnv_Level[#Level].Cnv2.Inputs.Lpd1;
   "HMI_CNV_Lpd2" := "Control_DB".LCnv_Sys[#System_No].Cnv_Level[#Level].Cnv2.Inputs.Lpd2;
   "HMI_CNV_Right" := "Control_DB".LCnv_Sys[#System_No].Cnv_Level[#Level].Cnv2.Inputs.Right;
   "HMI_CNV_Rpd1" := "Control_DB".LCnv_Sys[#System_No].Cnv_Level[#Level].Cnv2.Inputs.Rpd1;
   "HMI_CNV_Rpd2" := "Control_DB".LCnv_Sys[#System_No].Cnv_Level[#Level].Cnv2.Inputs.Rpd2;"HMI_CNV_Sdetect1" := "Control_DB".LCnv_Sys[#System_No].Cnv_Level[#Level].Cnv2.Inputs.Sdetect1;
   "HMI_CNV_Sdetect2" := "Control_DB".LCnv_Sys[#System_No].Cnv_Level[#Level].Cnv2.Inputs.Sdetect2;
   "HMI_CNV_SftyPinUp" := "Control_DB".LCnv_Sys[#System_No].Cnv_Level[#Level].Cnv2.Safety_Stop_Cnrl.Inputs.DP_Extended;
   "HMI_CNV_SftyPinDown" := "Control_DB".LCnv_Sys[#System_No].Cnv_Level[#Level].Cnv2.Safety_Stop_Cnrl.Inputs.DP_Retracted;
   IF "Control_DB".LCnv_Sys[#System_No].Cnv_Level[#Level].Cnv2.Safety_Stop_Cnrl.Inputs.DP_Extended AND
       NOT "Control_DB".LCnv_Sys[#System_No].Cnv_Level[#Level].Cnv2.Safety_Stop_Cnrl.Inputs.DP_Retracted THEN
       "UpDown" := 1;
   ELSIF NOT "Control_DB".LCnv_Sys[#System_No].Cnv_Level[#Level].Cnv2.Safety_Stop_Cnrl.Inputs.DP_Extended AND
       "Control_DB".LCnv_Sys[#System_No].Cnv_Level[#Level].Cnv2.Safety_Stop_Cnrl.Inputs.DP_Retracted THEN
       "UpDown" := 2;
   ELSE
       "UpDown" := 0;
   END_IF;

   //Feedback
   "Mode_HMI" := "Control_DB".LCnv_Sys[#System_No].Cnv_Level[#Level].Cnv2.Mode;
   "Enabled_HMI" := "Control_DB".LCnv_Sys[#System_No].Cnv_Level[#Level].Cnv2.Enabled;
   "Error_HMI" := "Control_DB".LCnv_Sys[#System_No].Cnv_Level[#Level].Cnv2.Error;
   "Warning_HMI" := "Control_DB".LCnv_Sys[#System_No].Cnv_Level[#Level].Cnv2.Warning;
   "Stopped_HMI" := "Control_DB".LCnv_Sys[#System_No].Cnv_Level[#Level].Cnv2.Stopped;
   "Running_HMI" := "Control_DB".LCnv_Sys[#System_No].Cnv_Level[#Level].Cnv2.Running;
   "Ready_For_Task_HMI" := "Control_DB".LCnv_Sys[#System_No].Cnv_Level[#Level].Cnv2.Ready_For_Task;
   "Cnv_Occupied_HMI" := "Control_DB".LCnv_Sys[#System_No].Cnv_Level[#Level].Cnv2.Cnv_Occupied;
   "Shuttle_in_place_HMI" := "Control_DB".LCnv_Sys[#System_No].Cnv_Level[#Level].Cnv2.Shuttle_In_Place;
   "Current_Task_Type_HMI" := "Control_DB".LCnv_Sys[#System_No].Cnv_Level[#Level].Cnv2.Current_Task_Type;
   "Current_Task_ID_HMI" := "Control_DB".LCnv_Sys[#System_No].Cnv_Level[#Level].Cnv2.Current_Task_ID;
   "SM_State_HMI" := "Control_DB".LCnv_Sys[#System_No].Cnv_Level[#Level].Cnv2.SM_State;
   IF "Control_DB".LCnv_Sys[#System_No].Cnv_Level[#Level].Cnv2.Motor.Forward THEN
       "Motor_Direction_HMI" := 1;
   ELSIF "Control_DB".LCnv_Sys[#System_No].Cnv_Level[#Level].Cnv2.Motor.Reverse THEN
       "Motor_Direction_HMI" := 2;
   ELSE
       "Motor_Direction_HMI" := 0;
   END_IF;
   "Motor_Speed_Requested_HMI" := "Control_DB".LCnv_Sys[#System_No].Cnv_Level[#Level].Cnv2.Motor.Speed;
   "Motor_Speed_Actual_HMI" := "Control_DB".LCnv_Sys[#System_No].Cnv_Level[#Level].Cnv2.Motor.Speed_Actual;
   "Transfer_To_ID_HMI" := "Control_DB".LCnv_Sys[#System_No].Cnv_Level[#Level].Cnv2.Instruction.Transfer_To_ID;
   "Transfer_From_ID_HMI" := "Control_DB".LCnv_Sys[#System_No].Cnv_Level[#Level].Cnv2.Instruction.Transfer_From_ID;

   //Instructions
   "Control_DB".LCnv_Sys[#System_No].Cnv_Level[#Level].Cnv2.Instruction.Stop := "Stop_HMI";
   "Control_DB".LCnv_Sys[#System_No].Cnv_Level[#Level].Cnv2.Instruction.Execute := "Manual_Fwd_HMI" OR "Manual_Bwd_HMI";
   "Control_DB".LCnv_Sys[#System_No].Cnv_Level[#Level].Cnv2.Instruction.Mode_Change := "Mode_Change_HMI";
   "Control_DB".LCnv_Sys[#System_No].Cnv_Level[#Level].Cnv2.Instruction.Enable := "Enable_HMI";
   "Control_DB".LCnv_Sys[#System_No].Cnv_Level[#Level].Cnv2.Instruction.Reset := "Reset_HMI";
   IF "Control_DB".LCnv_Sys[#System_No].Cnv_Level[#Level].Cnv2.Mode <> 3 THEN
       "Control_DB".LCnv_Sys[#System_No].Cnv_Level[#Level].Cnv2.Instruction.Foward := "Manual_Fwd_HMI";
       "Control_DB".LCnv_Sys[#System_No].Cnv_Level[#Level].Cnv2.Instruction.Backward := "Manual_Bwd_HMI";
       "Control_DB".LCnv_Sys[#System_No].Cnv_Level[#Level].Cnv2.Instruction.Start_Transfer := "Start_Transfer_HMI";
       IF "Control_DB".LCnv_Sys[#System_No].Cnv_Level[#Level].Cnv2.Mode = 1 THEN
           "Control_DB".LCnv_Sys[#System_No].Cnv_Level[#Level].Cnv2.Instruction.Start_Transfer_Backward := "Transfer_Backward";
       END_IF;
       "Control_DB".LCnv_Sys[#System_No].Cnv_Level[#Level].Cnv2.Safety_Stop_Cnrl.Instruction.Manual_Extend := "Manual_Sfty_Stopper_Up";
       "Control_DB".LCnv_Sys[#System_No].Cnv_Level[#Level].Cnv2.Safety_Stop_Cnrl.Instruction.Manual_Retract := "Manual_Sfty_Stopper_Down";
       "Control_DB".LCnv_Sys[#System_No].Cnv_Level[#Level].Cnv2.Instruction.Task_ID := "Task_ID_HMI";
       "Control_DB".LCnv_Sys[#System_No].Cnv_Level[#Level].Cnv2.Instruction.Pallet_Align_Left := "Pallet_Align_Left_HMI";
       "Control_DB".LCnv_Sys[#System_No].Cnv_Level[#Level].Cnv2.Instruction.Pallet_Align_Right := "Pallet_Align_Right_HMI";
       "Control_DB".LCnv_Sys[#System_No].Cnv_Level[#Level].Cnv2.Instruction.Pallet_Allignment := "Pallet_Align_Right_HMI";
       IF "CNV_HMI".In_Out[#System_No] THEN // 0 = Inbound, 1 = Outbound
           "Control_DB".LCnv_Sys[#System_No].Cnv_Level[#Level].Cnv2.Instruction.Transfer_To_ID := DINT#100000 + (#Level * 100) + #System_No;
           "Control_DB".LCnv_Sys[#System_No].Cnv_Level[#Level].Cnv2.Instruction.Transfer_From_ID := 0;
       ELSE
           "Control_DB".LCnv_Sys[#System_No].Cnv_Level[#Level].Cnv2.Instruction.Transfer_To_ID := 0;
           "Control_DB".LCnv_Sys[#System_No].Cnv_Level[#Level].Cnv2.Instruction.Transfer_From_ID := DINT#100000 + (#Level * 100+ #System_No);
       END_IF;
   END_IF;
END_FUNCTION

FUNCTION "Feed_ECNV(1)" : Void   // FC29, SCL
{ S7_Optimized_Access := 'TRUE' }
VERSION : 0.1
// stored: AutoNumber true, IsIECCheckEnabled false, SetENOAutomatically false, UDAEnableTagReadback false
   VAR_INPUT
      System_No : UInt;
   END_VAR
BEGIN
   //Sensors
   "HMI_CNV_Left(1)":= "Control_DB".ECnv_Sys[#System_No].Inputs.Left;
   "HMI_CNV_Lpd1(1)":= "Control_DB".ECnv_Sys[#System_No].Inputs.Lpd1;
   "HMI_CNV_Lpd2(1)":= "Control_DB".ECnv_Sys[#System_No].Inputs.Center;
   "HMI_CNV_Right(1)":= "Control_DB".ECnv_Sys[#System_No].Inputs.Right;
   "HMI_CNV_Rpd1(1)":= "Control_DB".ECnv_Sys[#System_No].Inputs.Rpd1;
   "HMI_CNV_Sdetect1(1)":= "Control_DB".ECnv_Sys[#System_No].Inputs.Overhang_Left;
   "HMI_CNV_Sdetect2(1)":= "Control_DB".ECnv_Sys[#System_No].Inputs.Overhang_Right;

   //Feedback
   "Mode_HMI(1)":= "Control_DB".ECnv_Sys[#System_No].Mode;
   "Enabled_HMI(1)":= "Control_DB".ECnv_Sys[#System_No].Enabled;
   "Error_HMI(1)":= "Control_DB".ECnv_Sys[#System_No].Error;
   "Warning_HMI(1)":= "Control_DB".ECnv_Sys[#System_No].Warning;
   "Stopped_HMI(1)":= "Control_DB".ECnv_Sys[#System_No].Stopped;
   "Running_HMI(1)":= "Control_DB".ECnv_Sys[#System_No].Running;
   "Ready_For_Task_HMI(1)":= "Control_DB".ECnv_Sys[#System_No].Ready_For_Task;
   "Cnv_Occupied_HMI(1)":= "Control_DB".ECnv_Sys[#System_No].Cnv_Occupied;
   "Shuttle_in_place_HMI(1)":= "Control_DB".ECnv_Sys[#System_No].Shuttle_In_Place;
   "Current_Task_Type_HMI(1)":= "Control_DB".ECnv_Sys[#System_No].Current_Task_Type;
   "Current_Task_ID_HMI(1)":= "Control_DB".ECnv_Sys[#System_No].Current_Task_ID;
   "SM_State_HMI(1)":= "Control_DB".ECnv_Sys[#System_No].SM_State;
   IF "Control_DB".ECnv_Sys[#System_No].Motor.Forward THEN
       "Motor_Direction_HMI(1)":= 1;
   ELSIF "Control_DB".ECnv_Sys[#System_No].Motor.Reverse THEN
       "Motor_Direction_HMI(1)":= 2;
   ELSE
       "Motor_Direction_HMI(1)":= 0;
   END_IF;
   "Motor_Speed_Requested_HMI(1)":= "Control_DB".ECnv_Sys[#System_No].Motor.Speed;
   "Motor_Speed_Actual_HMI(1)":= "Control_DB".ECnv_Sys[#System_No].Motor.Speed_Actual;
   "Transfer_To_ID_HMI(1)":= "Control_DB".ECnv_Sys[#System_No].Instruction.Transfer_To_ID;
   "Transfer_From_ID_HMI(1)":= "Control_DB".ECnv_Sys[#System_No].Instruction.Transfer_From_ID;

   //Instructions
   "Control_DB".ECnv_Sys[#System_No].Instruction.Stop := "Stop_HMI(1)";
   "Control_DB".ECnv_Sys[#System_No].Instruction.Execute := "Manual_Fwd_HMI(1)" OR "Manual_Bwd_HMI(1)";
   "Control_DB".ECnv_Sys[#System_No].Instruction.Mode_Change := "Mode_Change_HMI(1)";
   "Control_DB".ECnv_Sys[#System_No].Instruction.Enable := "Enable_HMI(1)";
   "Control_DB".ECnv_Sys[#System_No].Instruction.Reset := "Reset_HMI(1)";
   IF "Control_DB".ECnv_Sys[#System_No].Mode <> 3 THEN
       "Control_DB".ECnv_Sys[#System_No].Instruction.Foward := "Manual_Fwd_HMI(1)";
       "Control_DB".ECnv_Sys[#System_No].Instruction.Backward := "Manual_Bwd_HMI(1)";
       "Control_DB".ECnv_Sys[#System_No].Instruction.Start_Transfer := "Start_Transfer_HMI(1)";
       IF "Control_DB".ECnv_Sys[#System_No].Mode = 1 THEN
           "Control_DB".ECnv_Sys[#System_No].Instruction.Start_Transfer_Backward := "Transfer_Backward(1)";
       END_IF;
       "Control_DB".ECnv_Sys[#System_No].Instruction.Task_ID := "Task_ID_HMI(1)";
       "Control_DB".ECnv_Sys[#System_No].Instruction.Pallet_Align_Left := "Pallet_Align_Left_HMI(1)";
       "Control_DB".ECnv_Sys[#System_No].Instruction.Pallet_Align_Right := "Pallet_Align_Right_HMI(1)";
       "Control_DB".ECnv_Sys[#System_No].Instruction.Pallet_Allignment := "Pallet_Align_Right_HMI(1)";
       IF "CNV_HMI".In_Out[#System_No] THEN // 0 = Inbound, 1 = Outbound
           "Control_DB".ECnv_Sys[#System_No].Instruction.Transfer_To_ID := "CNV_ID_HMI(1)";
           "Control_DB".ECnv_Sys[#System_No].Instruction.Transfer_From_ID := 0;
       ELSE
           "Control_DB".ECnv_Sys[#System_No].Instruction.Transfer_To_ID := 0;
           "Control_DB".ECnv_Sys[#System_No].Instruction.Transfer_From_ID := "CNV_ID_HMI(1)";
       END_IF;
   END_IF;
END_FUNCTION

FUNCTION "Feed_ECNV" : Void   // FC1, SCL
{ S7_Optimized_Access := 'TRUE' }
VERSION : 0.1
// stored: AutoNumber true, IsIECCheckEnabled false, SetENOAutomatically false, UDAEnableTagReadback false
   VAR_INPUT
      System_No : UInt;
      Safety_OK : Bool;
      Overhang_Left : Bool;
      Overhang_Right : Bool;
   END_VAR
   VAR_IN_OUT
      System_Busy : Bool;
   END_VAR
BEGIN
   //Sensors
   "HMI_CNV_Left" := "Control_DB".ECnv_Sys[#System_No].Inputs.Left;
   "HMI_CNV_Lpd1" := "Control_DB".ECnv_Sys[#System_No].Inputs.Lpd1;
   "HMI_CNV_Lpd2" := "Control_DB".ECnv_Sys[#System_No].Inputs.Center;
   "HMI_CNV_Rpd1" := "Control_DB".ECnv_Sys[#System_No].Inputs.Rpd1;
   "HMI_CNV_Right" := "Control_DB".ECnv_Sys[#System_No].Inputs.Right;

   "HMI_CNV_Sdetect1" := #Overhang_Left;
   "HMI_CNV_Sdetect2" := #Overhang_Right;

   //Feedback
   "Mode_HMI" := "Control_DB".ECnv_Sys[#System_No].Mode;
   "Enabled_HMI" := "Control_DB".ECnv_Sys[#System_No].Enabled;
   "Error_HMI" := "Control_DB".ECnv_Sys[#System_No].Error;
   "Warning_HMI" := "Control_DB".ECnv_Sys[#System_No].Warning;
   "Stopped_HMI" := "Control_DB".ECnv_Sys[#System_No].Stopped;
   "Running_HMI" := "Control_DB".ECnv_Sys[#System_No].Running;
   "Ready_For_Task_HMI" := "Control_DB".ECnv_Sys[#System_No].Ready_For_Task;
   "Cnv_Occupied_HMI" := "Control_DB".ECnv_Sys[#System_No].Cnv_Occupied;
   "Shuttle_in_place_HMI" := "Control_DB".ECnv_Sys[#System_No].Shuttle_In_Place;
   "Current_Task_Type_HMI" := "Control_DB".ECnv_Sys[#System_No].Current_Task_Type;
   "Current_Task_ID_HMI" := "Control_DB".ECnv_Sys[#System_No].Current_Task_ID;
   "SM_State_HMI" := "Control_DB".ECnv_Sys[#System_No].SM_State;
   "Pallet_Type_HMI" := "Control_DB".ECnv_Sys[#System_No].Pallet_Type;
   IF "Control_DB".ECnv_Sys[#System_No].Motor.Forward THEN
       "Motor_Direction_HMI" := 1;
   ELSIF "Control_DB".ECnv_Sys[#System_No].Motor.Reverse THEN
       "Motor_Direction_HMI" := 2;
   ELSE
       "Motor_Direction_HMI" := 0;
   END_IF;
   "Motor_Speed_Requested_HMI" := "Control_DB".ECnv_Sys[#System_No].Motor.Speed;
   "Motor_Speed_Actual_HMI" := "Control_DB".ECnv_Sys[#System_No].Motor.Speed_Actual;
   "CNV_Motor_Ready" := "Control_DB".ECnv_Sys[#System_No].Motor.Ready;
   "CNV_Motor_Current_Actual_HMI" := "Control_DB".ECnv_Sys[#System_No].Motor.Actual_Current;
   "CNV_Motor_Actual_Torque" := "Control_DB".ECnv_Sys[#System_No].Motor.Actual_Torque;
   "Transfer_To_ID_HMI" := "Control_DB".ECnv_Sys[#System_No].Instruction.Transfer_To_ID;
   "Transfer_From_ID_HMI" := "Control_DB".ECnv_Sys[#System_No].Instruction.Transfer_From_ID;

   IF "Control_DB".ECnv_Sys[#System_No].Motor.Error THEN
       "CNV_Motor_Status_HMI" := 2;
   ELSIF "Control_DB".ECnv_Sys[#System_No].Motor.Enabled THEN
       "CNV_Motor_Status_HMI" := 1;
   ELSIF NOT "Control_DB".ECnv_Sys[#System_No].Motor.Enabled THEN
       "CNV_Motor_Status_HMI" := 0;
   END_IF;

   "Safety_OK_HMI" := #Safety_OK;

   //Instructions
   IF ("HMI_Box_Connected_1" = #System_No OR ("HMI_Box_Connected_1" >= (#System_No * 10) + 1 AND "HMI_Box_Connected_1" <= (#System_No * 10) + 8)) OR
       ("HMI_Box_Connected_2" = #System_No OR ("HMI_Box_Connected_1" >= (#System_No * 10) + 1 AND "HMI_Box_Connected_1" <= (#System_No * 10) + 8))
   THEN
       #System_Busy := TRUE;
   ELSE
       #System_Busy := FALSE;
       "Control_DB".ECnv_Sys[#System_No].Instruction.Stop := "Stop_HMI";
       "Control_DB".ECnv_Sys[#System_No].Instruction.Execute := "Manual_Fwd_HMI" OR "Manual_Bwd_HMI";
       IF "BT_Confirmation_HMI" THEN
           "Control_DB".VTD_Sys[#System_No].Instruction.Mode_Change :=
           "Control_DB".ECnv_Sys[#System_No].Instruction.Mode_Change :=
           "Control_DB".LCnv_Sys[#System_No].Cnv_Level[1].Cnv1.Instruction.Mode_Change :=
           "Control_DB".LCnv_Sys[#System_No].Cnv_Level[2].Cnv1.Instruction.Mode_Change :=
           "Control_DB".LCnv_Sys[#System_No].Cnv_Level[3].Cnv1.Instruction.Mode_Change :=
           "Control_DB".LCnv_Sys[#System_No].Cnv_Level[4].Cnv1.Instruction.Mode_Change :=
           "Control_DB".LCnv_Sys[#System_No].Cnv_Level[5].Cnv1.Instruction.Mode_Change :=
           "Control_DB".LCnv_Sys[#System_No].Cnv_Level[6].Cnv1.Instruction.Mode_Change :=
           "Control_DB".LCnv_Sys[#System_No].Cnv_Level[7].Cnv1.Instruction.Mode_Change :=
           "Control_DB".LCnv_Sys[#System_No].Cnv_Level[8].Cnv1.Instruction.Mode_Change :=
           "Control_DB".LCnv_Sys[#System_No].Cnv_Level[1].Cnv2.Instruction.Mode_Change :=
           "Control_DB".LCnv_Sys[#System_No].Cnv_Level[2].Cnv2.Instruction.Mode_Change :=
           "Control_DB".LCnv_Sys[#System_No].Cnv_Level[3].Cnv2.Instruction.Mode_Change :=
           "Control_DB".LCnv_Sys[#System_No].Cnv_Level[4].Cnv2.Instruction.Mode_Change :=
           "Control_DB".LCnv_Sys[#System_No].Cnv_Level[5].Cnv2.Instruction.Mode_Change :=
           "Control_DB".LCnv_Sys[#System_No].Cnv_Level[6].Cnv2.Instruction.Mode_Change :=
           "Control_DB".LCnv_Sys[#System_No].Cnv_Level[7].Cnv2.Instruction.Mode_Change :=
           "Control_DB".LCnv_Sys[#System_No].Cnv_Level[8].Cnv2.Instruction.Mode_Change := "Mode_Change_HMI";
           "Mode_Change_HMI(1)" := "Mode_Change_HMI";
           "BT_Confirmation_HMI" := FALSE;
       END_IF;

       "Control_DB".ECnv_Sys[#System_No].Instruction.Enable := "Enable_HMI";

       "Control_DB".ECnv_Sys[#System_No].Instruction.Reset := "Reset_HMI" OR "Reset_All" OR
       "Screen_DB_1".Reset_All[1] OR "CNV_HMI".Reset[1] OR
       "Screen_DB_1".Reset_All[2] OR "CNV_HMI".Reset[2];

       IF "Control_DB".ECnv_Sys[#System_No].Mode <> 3 THEN
           "Control_DB".ECnv_Sys[#System_No].Instruction.Foward := "Manual_Fwd_HMI";
           "Control_DB".ECnv_Sys[#System_No].Instruction.Backward := "Manual_Bwd_HMI";
           "Control_DB".ECnv_Sys[#System_No].Instruction.Start_Transfer := "Start_Transfer_HMI";
           IF "Control_DB".ECnv_Sys[#System_No].Mode = 1 THEN
               "Control_DB".ECnv_Sys[#System_No].Instruction.Start_Transfer_Backward := "Transfer_Backward";
           END_IF;
           "Control_DB".ECnv_Sys[#System_No].Instruction.Task_ID := "Task_ID_HMI";
           "Control_DB".ECnv_Sys[#System_No].Instruction.Pallet_Align_Left := "Pallet_Align_Left_HMI";
           "Control_DB".ECnv_Sys[#System_No].Instruction.Pallet_Align_Right := "Pallet_Align_Right_HMI";
           "Control_DB".ECnv_Sys[#System_No].Instruction.Pallet_Align_Center := "Pallet_Align_Center_HMI";
           IF "Mode_Change_HMI" <> 2 THEN
               "Control_DB".ECnv_Sys[#System_No].Instruction.Pallet_Allignment := "Pallet_Allignment_HMI" := FALSE;
           ELSE
               "Control_DB".ECnv_Sys[#System_No].Instruction.Pallet_Allignment := "Pallet_Allignment_HMI";
           END_IF;
           IF "CNV_HMI".In_Out[#System_No] THEN // 0 = ECNV RECEIVE, 1 = ECONV SEND
               "Control_DB".ECnv_Sys[#System_No].Instruction.Transfer_To_ID := "CNV_ID_HMI(1)";
               "Control_DB".ECnv_Sys[#System_No].Instruction.Transfer_From_ID := 0;
           ELSE
               "Control_DB".ECnv_Sys[#System_No].Instruction.Transfer_To_ID := 0;
               "Control_DB".ECnv_Sys[#System_No].Instruction.Transfer_From_ID := "CNV_ID_HMI(1)";
           END_IF;
       END_IF;
   END_IF;
END_FUNCTION

FUNCTION "Feed_ECNV_1" : Void   // FC53, SCL
{ S7_Optimized_Access := 'TRUE' }
VERSION : 0.1
// stored: AutoNumber true, IsIECCheckEnabled false, SetENOAutomatically false, UDAEnableTagReadback false
   VAR_INPUT
      HMI_No : UInt;
      HMI_Box : UInt;
      Overhang_Left : Bool;
      Overhang_Right : Bool;
      Sys_No : UInt;
      Safety_OK : Bool;
   END_VAR
BEGIN
   //Sensors
   "CNV_HMI".Left[#HMI_No] := "Control_DB".ECnv_Sys[#Sys_No].Inputs.Left;
   "CNV_HMI".Lpd1[#HMI_No] := "Control_DB".ECnv_Sys[#Sys_No].Inputs.Lpd1;
   "CNV_HMI".Center[#HMI_No] := "Control_DB".ECnv_Sys[#Sys_No].Inputs.Center;
   "CNV_HMI".Rpd1[#HMI_No] := "Control_DB".ECnv_Sys[#Sys_No].Inputs.Rpd1;
   "CNV_HMI".Right[#HMI_No] := "Control_DB".ECnv_Sys[#Sys_No].Inputs.Right;

   "CNV_HMI".Sdetect1[#HMI_No] := #Overhang_Left;
   "CNV_HMI".Sdetect2[#HMI_No] := #Overhang_Right;

   //Feedback
   "CNV_HMI".Mode[#HMI_No] := "Control_DB".ECnv_Sys[#Sys_No].Mode;
   "CNV_HMI".Enabled[#HMI_No] := "Control_DB".ECnv_Sys[#Sys_No].Enabled;
   "CNV_HMI".Error[#HMI_No] := "Control_DB".ECnv_Sys[#Sys_No].Error;
   "CNV_HMI".Warning[#HMI_No] := "Control_DB".ECnv_Sys[#Sys_No].Warning;
   "CNV_HMI".Stopped[#HMI_No] := "Control_DB".ECnv_Sys[#Sys_No].Stopped;
   "CNV_HMI".Running[#HMI_No] := "Control_DB".ECnv_Sys[#Sys_No].Running;
   "CNV_HMI".Ready_For_Task[#HMI_No] := "Control_DB".ECnv_Sys[#Sys_No].Ready_For_Task;
   "CNV_HMI".Occupied[#HMI_No] := "Control_DB".ECnv_Sys[#Sys_No].Cnv_Occupied;
   "CNV_HMI".Shuttle_in_place[#HMI_No] := "Control_DB".ECnv_Sys[#Sys_No].Shuttle_In_Place;
   "CNV_HMI".Current_Task_Type[#HMI_No] := "Control_DB".ECnv_Sys[#Sys_No].Current_Task_Type;
   "CNV_HMI".Current_Task_ID[#HMI_No] := "Control_DB".ECnv_Sys[#Sys_No].Current_Task_ID;
   "CNV_HMI".SM_State[#HMI_No] := "Control_DB".ECnv_Sys[#Sys_No].SM_State;
   "CNV_HMI".Pallet_Type[#HMI_No] := "Control_DB".ECnv_Sys[#Sys_No].Pallet_Type;
   IF "Control_DB".ECnv_Sys[#Sys_No].Motor.Forward THEN
       "CNV_HMI".Motor_Direction[#HMI_No] := 1;
   ELSIF "Control_DB".ECnv_Sys[#Sys_No].Motor.Reverse THEN
       "CNV_HMI".Motor_Direction[#HMI_No] := 2;
   ELSE
       "CNV_HMI".Motor_Direction[#HMI_No] := 0;
   END_IF;
   "CNV_HMI".Motor_Speed_Requested[#HMI_No] := "Control_DB".ECnv_Sys[#Sys_No].Motor.Speed;
   "CNV_HMI".Motor_Speed_Actual[#HMI_No] := "Control_DB".ECnv_Sys[#Sys_No].Motor.Speed_Actual;
   "CNV_HMI".Motor_Ready[#HMI_No] := "Control_DB".ECnv_Sys[#Sys_No].Motor.Ready;
   "CNV_HMI".Motor_Current_Actual[#HMI_No] := "Control_DB".ECnv_Sys[#Sys_No].Motor.Actual_Current;
   "CNV_HMI".Motor_Actual_Torque[#HMI_No] := "Control_DB".ECnv_Sys[#Sys_No].Motor.Actual_Torque;
   "CNV_HMI".Transfer_To_ID[#HMI_No] := "Control_DB".ECnv_Sys[#Sys_No].Instruction.Transfer_To_ID;
   "CNV_HMI".Transfer_From_ID[#HMI_No] := "Control_DB".ECnv_Sys[#Sys_No].Instruction.Transfer_From_ID;

   IF "Control_DB".ECnv_Sys[#Sys_No].Motor.Error THEN
       "CNV_HMI".Motor_Status[#HMI_No] := 2;
   ELSIF "Control_DB".ECnv_Sys[#Sys_No].Motor.Enabled THEN
       "CNV_HMI".Motor_Status[#HMI_No] := 1;
   ELSIF NOT "Control_DB".ECnv_Sys[#Sys_No].Motor.Enabled THEN
       "CNV_HMI".Motor_Status[#HMI_No] := 0;
   END_IF;

   "CNV_HMI".Safety_OK[#HMI_No] := #Safety_OK;

   //Instructions
   IF "Control_DB".VTD_Sys[#Sys_No].Current_Level = #HMI_Box MOD 10 THEN
       "Control_DB".ECnv_Sys[#Sys_No].Instruction.Stop := "CNV_HMI".Stop[#HMI_No];
       "Control_DB".ECnv_Sys[#Sys_No].Instruction.Execute := "CNV_HMI".Manual_Fwd[#HMI_No] OR "CNV_HMI".Manual_Bwd[#HMI_No];
       "Control_DB".ECnv_Sys[#Sys_No].Instruction.Mode_Change := "CNV_HMI".Mode_Change[#HMI_No];
       "Control_DB".ECnv_Sys[#Sys_No].Instruction.Enable := "CNV_HMI".Enable[#HMI_No];
       "Control_DB".ECnv_Sys[#Sys_No].Instruction.Reset := "CNV_HMI".Reset[#HMI_No] OR "Screen_DB_1".Reset_All[#HMI_No];
       IF "Control_DB".ECnv_Sys[#Sys_No].Mode <> 3 THEN
           "Control_DB".ECnv_Sys[#Sys_No].Instruction.Foward := "CNV_HMI".Manual_Fwd[#HMI_No];
           "Control_DB".ECnv_Sys[#Sys_No].Instruction.Backward := "CNV_HMI".Manual_Bwd[#HMI_No];
           "Control_DB".ECnv_Sys[#Sys_No].Instruction.Start_Transfer := "CNV_HMI".Start_Transfer[#HMI_No];
           "Control_DB".ECnv_Sys[#Sys_No].Instruction.Task_ID := "CNV_HMI".Task_ID[#HMI_No];
           "Control_DB".ECnv_Sys[#Sys_No].Instruction.Pallet_Align_Left := "CNV_HMI".Pallet_Align_Left[#HMI_No];
           "Control_DB".ECnv_Sys[#Sys_No].Instruction.Pallet_Align_Right := "CNV_HMI".Pallet_Align_Right[#HMI_No];
           "Control_DB".ECnv_Sys[#Sys_No].Instruction.Pallet_Align_Center := "CNV_HMI".Pallet_Align_Center[#HMI_No];
           IF "CNV_HMI".Mode_Change[#HMI_No] <> 2 THEN
               "Control_DB".ECnv_Sys[#Sys_No].Instruction.Pallet_Allignment := "CNV_HMI".Pallet_Allignment[#HMI_No] := FALSE;
           ELSE
               "Control_DB".ECnv_Sys[#Sys_No].Instruction.Pallet_Allignment := "CNV_HMI".Pallet_Allignment[#HMI_No];
           END_IF;
           IF "CNV_HMI".In_Out[#HMI_No] THEN // 0 = ECNV RECEIVE, 1 = ECONV SEND
               "Control_DB".ECnv_Sys[#Sys_No].Instruction.Transfer_To_ID := "CNV_HMI"."ID(1)"[#HMI_No];
               "Control_DB".ECnv_Sys[#Sys_No].Instruction.Transfer_From_ID := 0;
           ELSE
               "Control_DB".ECnv_Sys[#Sys_No].Instruction.Transfer_To_ID := 0;
               "Control_DB".ECnv_Sys[#Sys_No].Instruction.Transfer_From_ID := "CNV_HMI"."ID(1)"[#HMI_No];
           END_IF;
       END_IF;
   END_IF;
END_FUNCTION

FUNCTION "Feed_Steptable_FC" : Void   // FC44, SCL
{ S7_Optimized_Access := 'TRUE' }
VERSION : 0.1
// stored: AutoNumber true, IsIECCheckEnabled false, SetENOAutomatically false, UDAEnableTagReadback false
   VAR_INPUT
      CurrentTime : String;
      Task_Type : Int;
      Source_Location : DInt;
      Destination_Location : DInt;
      Pallet_Type : Char;
      Pallet_Alignment : Char;
      Shuttle_ID : Int;
   END_VAR
   VAR_IN_OUT
      StepTable : "OrderTable_UDT";
   END_VAR
BEGIN
   #StepTable.OrderNo := "OrderNo" + 1;
   #StepTable.StepNo := "OrderNo" + 1;
   #StepTable.PlaceTime := #CurrentTime;

   #StepTable.OPC_Control.Task_ID := "OrderNo" + 1;
   #StepTable.OPC_Control.Task_Type := #Task_Type;
   #StepTable.OPC_Control.Source_Location := #Source_Location;
   #StepTable.OPC_Control.Destination_Location := #Destination_Location;
   #StepTable.OPC_Control.Pallet_Type := #Pallet_Type;
   #StepTable.OPC_Control.Pallet_Alignment := #Pallet_Alignment;
   #StepTable.OPC_Control.Shuttle_ID := #Shuttle_ID;
END_FUNCTION

FUNCTION "Feed_VTD_HMI_FC" : Void   // FC33, SCL
{ S7_Optimized_Access := 'TRUE' }
VERSION : 0.1
// stored: AutoNumber true, IsIECCheckEnabled false, SetENOAutomatically false, UDAEnableTagReadback false
   VAR_INPUT
      Sys_No : UInt;
      Rem_Loc_Keys : Array[1..8] of Bool;
      Safety_OK : Bool;
      BCD_Test_Ok_HMI : Bool;
      BCD_Error_HMI : Bool;
      BCD_RdDone : Bool;
      BCD_ReqDone : Bool;
      BCD_ReqBusy : Bool;
      Start_InBarcodeStation : Bool;
      Sick_Lector_Reseult : String;
      Level_Below_Extractor : UInt;
      Speed_mm_s : Real;
   END_VAR
   VAR_OUTPUT
      System_Busy : Bool;
   END_VAR
   VAR_IN_OUT
      LE_Bypass : Bool;
      BCD_Start_Comm_Test_HMI : Bool;
      BCD_Enable_Trigger_HMI : Bool;
      BCD_Disable_Trigger_HMI : Bool;
      BCD_Execute_Function : Bool;
   END_VAR
BEGIN
   //Status
   "VTD_Error_HMI" := "Control_DB".VTD_Sys[#Sys_No].Error;
   "VTD_Warning_HMI" := "Control_DB".VTD_Sys[#Sys_No].Warning <> 0;
   "VTD_Enabled_HMI" := "Control_DB".VTD_Sys[#Sys_No].Enabled;
   "VTD_Stopped_HMI" := "Control_DB".VTD_Sys[#Sys_No].Stopped;
   "VTD_Running_HMI" := "Control_DB".VTD_Sys[#Sys_No].Running;
   "VTD_Docked_HMI" := "Control_DB".VTD_Sys[#Sys_No].Docked;
   "Safety_OK_HMI" := #Safety_OK;
   "VTD_Current_Task_Type_HMI" := "Control_DB".VTD_Sys[#Sys_No].Current_Task_Type;
   "VTD_Current_Task_ID_HMI" := "Control_DB".VTD_Sys[#Sys_No].Current_Task_ID;
   "VTD_Current_Level_HMI" := "Control_DB".VTD_Sys[#Sys_No].Current_Level;
   "VTD_LP_State_HMI" := "Control_DB".VTD_Sys[#Sys_No].LP_State;
   "VTD_Pallet_Type_HMI" := "Control_DB".VTD_Sys[#Sys_No].Pallet_Loaded;
   "VTD_Shuttle_Loaded_HMI" := "Control_DB".VTD_Sys[#Sys_No].Shuttle_Loaded;
   "VTD_SM_State_HMI" := "Control_DB".VTD_Sys[#Sys_No].SM_State;
   "VTD_LE_Error_HMI" := "Control_DB".VTD_Sys[#Sys_No].Inputs.LE_Status.%X0;
   "VTD_AE_Error_HMI" := "Control_DB".VTD_Sys[#Sys_No].Inputs.AE_Status_2.%X15;
   "VTD_Encoder_Delta_HMI" := "Control_DB".VTD_Sys[#Sys_No].Encoder_Delta;
   "VTD_Moving_To_Level" := "Control_DB".VTD_Sys[#Sys_No].Instruction.Move_To_Level;
   "VTD_Cnv_Occupied" := "Control_DB".VTD_Sys[#Sys_No].Pallet_Loaded <> 0;
   "VTD_Progress_HMI" := REAL_TO_INT("Control_DB".VTD_Sys[#Sys_No].LE);
   "VTD_Motor_SetPoint_HMI" := "Control_DB".VTD_Sys[#Sys_No].Motor_Speed;
   "VTD_Motor_Actual_Speed_HMI" := INT_TO_UINT("Control_DB".VTD_Sys[#Sys_No].Motor.Speed_Actual);
   "VTD_Motor_Actual_Current_HMI" := "Control_DB".VTD_Sys[#Sys_No].Motor.Actual_Current;
   "VTD_Actual_Torque" := "Control_DB".VTD_Sys[#Sys_No].Motor.Actual_Torque;
   "VTD_Motor_Ready_HMI" := "Control_DB".VTD_Sys[#Sys_No].Motor.Ready;
   "VTD_Level_Below_Extractor" := #Level_Below_Extractor;
   "VTD_Speed_mm_s" := #Speed_mm_s;
   "VTD_Mode_HMI" := "Control_DB".VTD_Sys[#Sys_No].Mode;

   //MOTOR STATUS
   IF "Control_DB".VTD_Sys[#Sys_No].Motor.Error THEN
       "VTD_Motor_Status_HMI" := 2;
   ELSIF "Control_DB".VTD_Sys[#Sys_No].Motor.Enabled THEN
       "VTD_Motor_Status_HMI" := 1;
   ELSIF NOT "Control_DB".VTD_Sys[#Sys_No].Motor.Enabled THEN
       "VTD_Motor_Status_HMI" := 0;
   END_IF;

   //BARCODE
   "BCD_Test_Ok_HMI" := #BCD_Test_Ok_HMI;
   "BCD_Error_HMI" := #BCD_Error_HMI;
   "BCD_RdDone" := #BCD_RdDone;
   "BCD_ReqDone" := #BCD_ReqDone;
   "BCD_ReqBusy" := #BCD_ReqBusy;
   "PopUps_DB".Sick_Lector_Reseult := #Sick_Lector_Reseult;

   //Inputs
   "VTD_Upper_Overtravel_HMI" := "Control_DB".VTD_Sys[#Sys_No].Inputs.Upper_Overtravel;
   "VTD_Upper_Limet_HMI" := "Control_DB".VTD_Sys[#Sys_No].Inputs.Upper_limit;
   "VTD_Ultimate_Slow_HMI" := "Control_DB".VTD_Sys[#Sys_No].Inputs.Ultimate_SlowDown;
   "VTD_Ultimate_Creep_HMI" := "Control_DB".VTD_Sys[#Sys_No].Inputs.Ultimate_Creep;
   "VTD_Lower_Limit_HMI" := "Control_DB".VTD_Sys[#Sys_No].Inputs.Lower_Limit;
   "VTD_Lower_Overtravel_HMI" := "Control_DB".VTD_Sys[#Sys_No].Inputs.Lower_Overtravel;
   "VTD_Level_Detect1_HMI" := "Control_DB".VTD_Sys[#Sys_No].Inputs.Level_Detect1;
   "VTD_Level_Detect2_HMI" := "Control_DB".VTD_Sys[#Sys_No].Inputs.Level_Detect2;
   "VTD_Ultimate_Slow_HMI" := "Control_DB".VTD_Sys[#Sys_No].Inputs.Ultimate_SlowDown;
   "VTD_Ultimate_Creep_HMI" := "Control_DB".VTD_Sys[#Sys_No].Inputs.Ultimate_Creep;
   "VTD_DP1_Extended_HMI" := "Control_DB".VTD_Sys[#Sys_No].Inputs.DP1_Extended;
   "VTD_DP2_Extended_HMI" := "Control_DB".VTD_Sys[#Sys_No].Inputs.DP2_Extended;
   "VTD_DP1_Retracted_HMI" := "Control_DB".VTD_Sys[#Sys_No].Inputs.DP1_Retracted;
   "VTD_DP2_Retracted_HMI" := "Control_DB".VTD_Sys[#Sys_No].Inputs.DP2_Retracted;
   "Chain Slack 1" := NOT "Control_DB".VTD_Sys[#Sys_No].Inputs.Chain_Slack_1;
   "Chain Slack 2" := NOT "Control_DB".VTD_Sys[#Sys_No].Inputs.Chain_Slack_2;
   "Chain Slack 3" := NOT "Control_DB".VTD_Sys[#Sys_No].Inputs.Chain_Slack_3;
   "Chain Slack 4" := NOT "Control_DB".VTD_Sys[#Sys_No].Inputs.Chain_Slack_4;
   "VTD_AE_HMI" := "Control_DB".VTD_Sys[#Sys_No].AE;
   "VTD_LE_HMI" := "Control_DB".VTD_Sys[#Sys_No].LE;
   "VTD_LE_Speed_HMI" := "Control_DB".VTD_Sys[#Sys_No].Inputs.LE_Speed;
   "LE_X_Unsafe_Position" := "Control_DB".VTD_Sys[#Sys_No].Inputs.LE_Position;
   "LE_Speed" := "Control_DB".VTD_Sys[#Sys_No].Inputs.LE_Speed;
   "LE_Warnings" := "Control_DB".VTD_Sys[#Sys_No].Inputs.LE_Warnings;
   "LE_Quality_Decoded_Codes" := "Control_DB".VTD_Sys[#Sys_No].Inputs.LE_Quality_Decoded_Codes;
   "LE_Quality_Value" := "Control_DB".VTD_Sys[#Sys_No].Inputs.LE_Quality_Value;

   "AE_Position_1" := "Control_DB".VTD_Sys[#Sys_No].Inputs.AE_Position_1;
   "AE_Position_2" := "Control_DB".VTD_Sys[#Sys_No].Inputs.AE_Position_2;
   "AE_Speed" := "Control_DB".VTD_Sys[#Sys_No].Inputs.AE_Speed;
   "AE_Status_1" := "Control_DB".VTD_Sys[#Sys_No].Inputs.AE_Status_1;
   "AE_Status_2" := "Control_DB".VTD_Sys[#Sys_No].Inputs.AE_Status_2;

   //Instruction
   IF "HMI_Box_Connected_1" <> 0 THEN
       IF "HMI_Box_Connected_1" = (#Sys_No * 10) + 9 OR
           ("HMI_Box_Connected_1" = (#Sys_No * 10) + "HMI_Box_Connected_1" MOD 10 AND #Rem_Loc_Keys["HMI_Box_Connected_1" MOD 10])
       THEN
           #System_Busy := TRUE;
       END_IF;
   END_IF;
   IF "HMI_Box_Connected_2" <> 0 THEN
       IF "HMI_Box_Connected_2" = (#Sys_No * 10) + 9 OR
           ("HMI_Box_Connected_2" = (#Sys_No * 10) + "HMI_Box_Connected_2" MOD 10 AND #Rem_Loc_Keys["HMI_Box_Connected_2" MOD 10])
       THEN
           #System_Busy := TRUE;
       END_IF;
   END_IF;

   IF NOT #System_Busy THEN
       #System_Busy := FALSE;
       IF NOT "Screen_DB".Charge_VTD_Commands THEN
           "Control_DB".VTD_Sys[#Sys_No].Instruction.Reset := "VTD_Reset_HMIs" OR "Reset_All" OR "VTD_HMI".Reset[1] OR "VTD_HMI".Reset[2] OR "Screen_DB_1".Reset_All[1] OR "Screen_DB_1".Reset_All[2];
           IF "BT_Confirmation_HMI" THEN
               "Control_DB".VTD_Sys[#Sys_No].Instruction.Mode_Change :=
               "Control_DB".ECnv_Sys[#Sys_No].Instruction.Mode_Change :=
               "Control_DB".LCnv_Sys[#Sys_No].Cnv_Level[1].Cnv1.Instruction.Mode_Change :=
               "Control_DB".LCnv_Sys[#Sys_No].Cnv_Level[2].Cnv1.Instruction.Mode_Change :=
               "Control_DB".LCnv_Sys[#Sys_No].Cnv_Level[3].Cnv1.Instruction.Mode_Change :=
               "Control_DB".LCnv_Sys[#Sys_No].Cnv_Level[4].Cnv1.Instruction.Mode_Change :=
               "Control_DB".LCnv_Sys[#Sys_No].Cnv_Level[5].Cnv1.Instruction.Mode_Change :=
               "Control_DB".LCnv_Sys[#Sys_No].Cnv_Level[6].Cnv1.Instruction.Mode_Change :=
               "Control_DB".LCnv_Sys[#Sys_No].Cnv_Level[7].Cnv1.Instruction.Mode_Change :=
               "Control_DB".LCnv_Sys[#Sys_No].Cnv_Level[8].Cnv1.Instruction.Mode_Change :=
               "Control_DB".LCnv_Sys[#Sys_No].Cnv_Level[1].Cnv2.Instruction.Mode_Change :=
               "Control_DB".LCnv_Sys[#Sys_No].Cnv_Level[2].Cnv2.Instruction.Mode_Change :=
               "Control_DB".LCnv_Sys[#Sys_No].Cnv_Level[3].Cnv2.Instruction.Mode_Change :=
               "Control_DB".LCnv_Sys[#Sys_No].Cnv_Level[4].Cnv2.Instruction.Mode_Change :=
               "Control_DB".LCnv_Sys[#Sys_No].Cnv_Level[5].Cnv2.Instruction.Mode_Change :=
               "Control_DB".LCnv_Sys[#Sys_No].Cnv_Level[6].Cnv2.Instruction.Mode_Change :=
               "Control_DB".LCnv_Sys[#Sys_No].Cnv_Level[7].Cnv2.Instruction.Mode_Change :=
               "Control_DB".LCnv_Sys[#Sys_No].Cnv_Level[8].Cnv2.Instruction.Mode_Change := "VTD_Mode_Change_HMI";
               "Control_DB".VTD_Sys[#Sys_No].Instruction.Move_To_Level := "VTD_Move_To_Level_HMI";
               "VTD_Move_To_Level_HMI" := 0;
               "BT_Confirmation_HMI" := FALSE;
           END_IF;

           "Control_DB".VTD_Sys[#Sys_No].Instruction.Enable := "VTD_Enable_HMI";
           IF "VTD_Stop_HMI" THEN
               "Control_DB".VTD_Sys[#Sys_No].Instruction.Stop := TRUE;
           END_IF;

           IF "Reset_All" OR "VTD_Reset_HMIs"
           THEN
               "Control_DB".VTD_Sys[#Sys_No].Instruction.Stop := "VTD_Stop_HMI" := FALSE;
           END_IF;

           IF "Control_DB".VTD_Sys[#Sys_No].Mode <> 3 THEN
               "Control_DB".VTD_Sys[#Sys_No].Instruction.Pallet_Type := "VTD_Pallet_Type_HMI";
               "Control_DB".VTD_Sys[#Sys_No].Instruction.Task_ID := "VTD_Task_ID_HMI";

               // IF "Control_DB".VTD_Sys[#Sys_No].Mode = 2 AND "VTD_Move_To_Level_HMI" <> 0 AND "BT_Confirmation_HMI" THEN
               //     "Control_DB".VTD_Sys[#Sys_No].Instruction.Move_To_Level := "VTD_Move_To_Level_HMI";
               //     "VTD_Move_To_Level_HMI" := 0;
               //     "BT_Confirmation_HMI" := 0;
               // END_IF;

               "Control_DB".VTD_Sys[#Sys_No].Instruction.Manual_Up := "VTD_Manual_Up_HMI";
               "Control_DB".VTD_Sys[#Sys_No].Instruction.Manual_Down := "VTD_Manual_Down_HMI";
               "Control_DB".VTD_Sys[#Sys_No].Instruction.Manual_LP_Retract := "VTD_Manual_LP_Retract_HMIs";
               "Control_DB".VTD_Sys[#Sys_No].Instruction.Manual_LP_Extend := "VTD_Manual_LP_Extend_HMIs";
               "Control_DB".VTD_Sys[#Sys_No].Instruction.Start_Teach := "VTD_Start_Teach_HMIs";
           END_IF;

           //ABSOLUTE ENCODER
           "Control_DB".VTD_Sys[#Sys_No].Outputs.AE_Control_Word_1 := "AE_Control_Word_1";
           "Control_DB".VTD_Sys[#Sys_No].Outputs.AE_Control_Word_2 := "AE_Control_Word_2";

           //LINEAR ENCODER
           #LE_Bypass := "LE_Bypass";

           IF "Control_DB".VTD_Sys[#Sys_No].LE > 0 THEN
               "LE_Bypass" := FALSE;
           END_IF;

           //BARCODE
           #BCD_Start_Comm_Test_HMI := "BCD_Start_Comm_Test_HMI";
           #BCD_Enable_Trigger_HMI := "BCD_Enable_Trigger_HMI";
           #BCD_Disable_Trigger_HMI := "BCD_Disable_Trigger_HMI";
           #BCD_Execute_Function := "BCD_Execute_Function";

           //SICK BARCODE MANUAL TRIG FROM HMI
           IF "Control_DB".VTD_Sys[#Sys_No].Mode <> 3 THEN
               "Control_DB".VTDBarcode_Station[#Sys_No].Start := #Start_InBarcodeStation;
           END_IF;
       END_IF;
   END_IF;
END_FUNCTION

FUNCTION "Feed_VTD_HMI_FC_1" : Void   // FC57, SCL
{ S7_Optimized_Access := 'TRUE' }
VERSION : 0.1
// stored: AutoNumber true, IsIECCheckEnabled false, SetENOAutomatically false, UDAEnableTagReadback false
   VAR_INPUT
      HMI_No : UInt;
      HMI_Box : UInt;
      Sys_No : UInt;
      Safety_OK : Bool;
      BCD_Test_Ok_HMI : Bool;
      BCD_Error_HMI : Bool;
      BCD_RdDone : Bool;
      BCD_ReqDone : Bool;
      BCD_ReqBusy : Bool;
      Sick_Lector_Reseult : String;
      Level_Below_Extractor : UInt;
      Speed_mm_s : Real;
   END_VAR
   VAR_IN_OUT
      BCD_Start_Comm_Test_HMI : Bool;
      BCD_Enable_Trigger_HMI : Bool;
      BCD_Disable_Trigger_HMI : Bool;
      BCD_Execute_Function : Bool;
   END_VAR
BEGIN
   //Status
   "VTD_HMI".Error[#HMI_No] := "Control_DB".VTD_Sys[#Sys_No].Error;
   "VTD_HMI".Warning[#HMI_No] := "Control_DB".VTD_Sys[#Sys_No].Warning <> 0;
   "VTD_HMI".Enabled[#HMI_No] := "Control_DB".VTD_Sys[#Sys_No].Enabled;
   "VTD_HMI".Stopped[#HMI_No] := "Control_DB".VTD_Sys[#Sys_No].Stopped;
   "VTD_HMI".Running[#HMI_No] := "Control_DB".VTD_Sys[#Sys_No].Running;
   "VTD_HMI".Docked[#HMI_No] := "Control_DB".VTD_Sys[#Sys_No].Docked;
   "VTD_HMI".Safety_OK[#HMI_No] := #Safety_OK;
   "VTD_HMI".Current_Task_Type[#HMI_No] :="Control_DB".VTD_Sys[#Sys_No].Current_Task_Type;
   "VTD_HMI".Current_Task_ID[#HMI_No] := "Control_DB".VTD_Sys[#Sys_No].Current_Task_ID;
   "VTD_HMI".Current_Level[#HMI_No] := "Control_DB".VTD_Sys[#Sys_No].Current_Level;
   "VTD_HMI".DP_State[#HMI_No] := "Control_DB".VTD_Sys[#Sys_No].LP_State;
   "VTD_HMI".Pallet_Type[#HMI_No] := "Control_DB".VTD_Sys[#Sys_No].Pallet_Loaded;
   "VTD_HMI".Shuttle_Loaded[#HMI_No] := "Control_DB".VTD_Sys[#Sys_No].Shuttle_Loaded;
   "VTD_HMI".SM_State[#HMI_No] := "Control_DB".VTD_Sys[#Sys_No].SM_State;
   "VTD_HMI".LE_Error[#HMI_No] := "Control_DB".VTD_Sys[#Sys_No].Inputs.LE_Status.%X0;
   "VTD_HMI".AE_Error[#HMI_No] := "Control_DB".VTD_Sys[#Sys_No].Inputs.AE_Status_2.%X15;
   "VTD_HMI".Encoder_Delta[#HMI_No] := "Control_DB".VTD_Sys[#Sys_No].Encoder_Delta;
   "VTD_HMI".Moving_To_Level[#HMI_No] := "Control_DB".VTD_Sys[#Sys_No].Instruction.Move_To_Level;
   "VTD_HMI".Cnv_Occupied[#HMI_No] := "Control_DB".VTD_Sys[#Sys_No].Pallet_Loaded <> 0;
   "VTD_HMI".Progress[#HMI_No] := REAL_TO_INT("Control_DB".VTD_Sys[#Sys_No].LE);
   "VTD_HMI".Motor_SetPoint[#HMI_No] := "Control_DB".VTD_Sys[#Sys_No].Motor_Speed;
   "VTD_HMI".Motor_Actual_Speed[#HMI_No] := INT_TO_UINT("Control_DB".VTD_Sys[#Sys_No].Motor.Speed_Actual);
   "VTD_HMI".Motor_Actual_Current[#HMI_No] := "Control_DB".VTD_Sys[#Sys_No].Motor.Actual_Current;
   "VTD_HMI".Actual_Torque[#HMI_No] := "Control_DB".VTD_Sys[#Sys_No].Motor.Actual_Torque;
   "VTD_HMI".Motor_Ready[#HMI_No] := "Control_DB".VTD_Sys[#Sys_No].Motor.Ready;
   "VTD_HMI".Level_Below_Extractor[#HMI_No] := #Level_Below_Extractor;
   "VTD_HMI".Speed_mm_s[#HMI_No] := #Speed_mm_s;
   "VTD_Mode_HMI" := "Control_DB".VTD_Sys[#Sys_No].Mode;

   //MOTOR STATUS
   IF "Control_DB".VTD_Sys[#Sys_No].Motor.Error THEN
       "VTD_HMI".Motor_Status[#HMI_No] := 2;
   ELSIF "Control_DB".VTD_Sys[#Sys_No].Motor.Enabled THEN
       "VTD_HMI".Motor_Status[#HMI_No] := 1;
   ELSIF NOT "Control_DB".VTD_Sys[#Sys_No].Motor.Enabled THEN
       "VTD_HMI".Motor_Status[#HMI_No] := 0;
   END_IF;

   //BARCODE
   "PopUps_DB_1".Lector_Barcode[#HMI_No].BCD_Test_Ok := #BCD_Test_Ok_HMI;
   "PopUps_DB_1".Lector_Barcode[#HMI_No].BCD_Error := #BCD_Error_HMI;
   "PopUps_DB_1".Lector_Barcode[#HMI_No].BCD_RdDone := #BCD_RdDone;
   "PopUps_DB_1".Lector_Barcode[#HMI_No].BCD_ReqDone := #BCD_ReqDone;
   "PopUps_DB_1".Lector_Barcode[#HMI_No].BCD_ReqBusy := #BCD_ReqBusy;
   "PopUps_DB_1".Lector_Barcode[#HMI_No].Lector_Reseult := #Sick_Lector_Reseult;

   //Inputs
   "VTD_HMI".Upper_Overtravel[#HMI_No] := "Control_DB".VTD_Sys[#Sys_No].Inputs.Upper_Overtravel;
   "VTD_HMI".Upper_Limet[#HMI_No] := "Control_DB".VTD_Sys[#Sys_No].Inputs.Upper_limit;
   "VTD_HMI".Ultimate_Slow[#HMI_No] := "Control_DB".VTD_Sys[#Sys_No].Inputs.Ultimate_SlowDown;
   "VTD_HMI".Ultimate_Creep[#Sys_No] := "Control_DB".VTD_Sys[#Sys_No].Inputs.Ultimate_Creep;
   "VTD_HMI".Lower_Limit[#HMI_No] := "Control_DB".VTD_Sys[#Sys_No].Inputs.Lower_Limit;
   "VTD_HMI".Lower_Overtravel[#HMI_No] := "Control_DB".VTD_Sys[#Sys_No].Inputs.Lower_Overtravel;
   "VTD_HMI".Level_Detect1[#HMI_No] := "Control_DB".VTD_Sys[#Sys_No].Inputs.Level_Detect1;
   "VTD_HMI".Level_Detect2[#HMI_No] := "Control_DB".VTD_Sys[#Sys_No].Inputs.Level_Detect2;
   "VTD_HMI".DP1_Extended[#HMI_No] := "Control_DB".VTD_Sys[#Sys_No].Inputs.DP1_Extended;
   "VTD_HMI".DP2_Extended[#HMI_No] := "Control_DB".VTD_Sys[#Sys_No].Inputs.DP2_Extended;
   "VTD_HMI".DP1_Retracted[#HMI_No] := "Control_DB".VTD_Sys[#Sys_No].Inputs.DP1_Retracted;
   "VTD_HMI".DP2_Retracted[#HMI_No] := "Control_DB".VTD_Sys[#Sys_No].Inputs.DP2_Retracted;
   "VTD_HMI"."Chain Slack 1"[#HMI_No] := NOT "Control_DB".VTD_Sys[#Sys_No].Inputs.Chain_Slack_1;
   "VTD_HMI"."Chain Slack 2"[#HMI_No] := NOT "Control_DB".VTD_Sys[#Sys_No].Inputs.Chain_Slack_2;
   "VTD_HMI"."Chain Slack 3"[#HMI_No] := NOT "Control_DB".VTD_Sys[#Sys_No].Inputs.Chain_Slack_3;
   "VTD_HMI"."Chain Slack 4"[#HMI_No] := NOT "Control_DB".VTD_Sys[#Sys_No].Inputs.Chain_Slack_4;
   "VTD_HMI".AE[#HMI_No] := "Control_DB".VTD_Sys[#Sys_No].AE;
   "VTD_HMI".LE[#HMI_No] := "Control_DB".VTD_Sys[#Sys_No].LE;
   "PopUps_DB_1".Linear_Encoder[#HMI_No].LE_Speed := "Control_DB".VTD_Sys[#Sys_No].Inputs.LE_Speed;
   "PopUps_DB_1".Linear_Encoder[#HMI_No].LE_X_Unsafe_Position := "Control_DB".VTD_Sys[#Sys_No].Inputs.LE_Position;
   "PopUps_DB_1".Linear_Encoder[#HMI_No].LE_Speed := "Control_DB".VTD_Sys[#Sys_No].Inputs.LE_Speed;
   "PopUps_DB_1".Linear_Encoder[#HMI_No].LE_Warnings := "Control_DB".VTD_Sys[#Sys_No].Inputs.LE_Warnings;

